// TwinCAT 3 PLC project Tc3UnitTest
// Title: Tc3_UnitTest
// Company: Lorenz Software
// ProjectVersion: 1.0.0.0
// ProgramVersion: 3.1.4026.27
// libraries:
//   Tc2_Standard, * (Beckhoff Automation GmbH)
//   Tc2_System, * (Beckhoff Automation GmbH)
//   Tc2_Utilities, * (Beckhoff Automation GmbH)
// project tree:
//   Framework/Assertions/DataTypes/ AssertionLRealRepresentation.TcDUT, AssertionRealRepresentation.TcDUT
//   Framework/Assertions/GlobalVariables/ Param_Assertions.TcGVL
//   Framework/Assertions/Interfaces/ I_Assertion.TcIO
//   Framework/Assertions/POU/Arrays/Bool/ AssertArrayAllEqual_Bool.TcPOU, AssertArrayContainsArray_Bool.TcPOU, AssertArrayContainsValue_Bool.TcPOU, AssertArrayNoValueChange_Bool.TcPOU, AssertEqualArray_Bool.TcPOU
//   Framework/Assertions/POU/Arrays/Byte/ AssertArrayAllEqual_Byte.TcPOU, AssertArrayContainsArray_Byte.TcPOU, AssertArrayContainsString_Byte.TcPOU, AssertArrayContainsValue_Byte.TcPOU, AssertArrayEndsWithArray_Byte.TcPOU, AssertArrayEndsWithString_Byte.TcPOU, AssertArrayEqualString_Byte.TcPOU, AssertArrayNoValueChange_Byte.TcPOU, AssertArrayStartsWithArray_Byte.TcPOU, AssertArrayStartsWithString_Byte.TcPOU, AssertEqualArray_Byte.TcPOU
//   Framework/Assertions/POU/Arrays/Byte/LengthUntilToken/ AssertLengthUntilArrayEqual_Byte.TcPOU (not stored), AssertLengthUntilArrayGreaterEqual_Byte.TcPOU (not stored), AssertLengthUntilArrayGreaterThan_Byte.TcPOU (not stored), AssertLengthUntilArrayLessEqual_Byte.TcPOU (not stored), AssertLengthUntilArrayLessThan_Byte.TcPOU (not stored), AssertLengthUntilArrayNotEqual_Byte.TcPOU (not stored), AssertLengthUntilValueEqual_Byte.TcPOU (not stored), AssertLengthUntilValueGreaterEqual_Byte.TcPOU (not stored), AssertLengthUntilValueGreaterThan_Byte.TcPOU (not stored), AssertLengthUntilValueLessEqual_Byte.TcPOU (not stored), AssertLengthUntilValueLessThan_Byte.TcPOU (not stored), AssertLengthUntilValueNotEqual_Byte.TcPOU (not stored)
//   Framework/Assertions/POU/Arrays/Byte/TokenCount/ AssertArrayTokenCntEqual_Byte.TcPOU (not stored), AssertArrayTokenCntGreaterEqual_Byte.TcPOU (not stored), AssertArrayTokenCntGreaterThan_Byte.TcPOU (not stored), AssertArrayTokenCntInRange_Byte.TcPOU (not stored), AssertArrayTokenCntLessEqual_Byte.TcPOU (not stored), AssertArrayTokenCntLessThan_Byte.TcPOU (not stored), AssertArrayTokenCntNotEqual_Byte.TcPOU (not stored), AssertArrayTokenCntNotInRange_Byte.TcPOU (not stored), AssertNoArrayToken_Byte.TcPOU (not stored), AssertNoValueToken_Byte.TcPOU (not stored), AssertValueTokenCntEqual_Byte.TcPOU (not stored), AssertValueTokenCntGreaterEqual_Byte.TcPOU (not stored), AssertValueTokenCntGreaterThan_Byte.TcPOU (not stored), AssertValueTokenCntInRange_Byte.TcPOU (not stored), AssertValueTokenCntLessEqual_Byte.TcPOU (not stored), AssertValueTokenCntLessThan_Byte.TcPOU (not stored), AssertValueTokenCntNotEqual_Byte.TcPOU (not stored), AssertValueTokenCntNotInRange_Byte.TcPOU (not stored)
//   Framework/Assertions/POU/Arrays/Char/ AssertArrayAllEqual_Char.TcPOU, AssertArrayContainsArray_Char.TcPOU, AssertArrayContainsString_Char.TcPOU, AssertArrayContainsValue_Char.TcPOU, AssertArrayEndsWithString_Char.TcPOU, AssertArrayEqualString_Char.TcPOU, AssertArrayNoValueChange_Char.TcPOU, AssertArrayStartsWithString_Char.TcPOU, AssertEqualArray_Char.TcPOU
//   Framework/Assertions/POU/Arrays/DInt/ AssertArrayAllEqual_DInt.TcPOU, AssertArrayContainsArray_DInt.TcPOU, AssertArrayContainsValue_DInt.TcPOU, AssertArrayNoValueChange_DInt.TcPOU, AssertEqualArray_DInt.TcPOU
//   Framework/Assertions/POU/Arrays/DWord/ AssertArrayAllEqual_DWord.TcPOU, AssertArrayContainsArray_DWord.TcPOU, AssertArrayContainsValue_DWord.TcPOU, AssertArrayNoValueChange_DWord.TcPOU, AssertEqualArray_DWord.TcPOU
//   Framework/Assertions/POU/Arrays/Int/ AssertArrayAllEqual_Int.TcPOU, AssertArrayContainsArray_Int.TcPOU, AssertArrayContainsValue_Int.TcPOU, AssertArrayNoValueChange_Int.TcPOU, AssertEqualArray_Int.TcPOU
//   Framework/Assertions/POU/Arrays/LInt/ AssertArrayAllEqual_LInt.TcPOU, AssertArrayContainsArray_LInt.TcPOU, AssertArrayContainsValue_LInt.TcPOU, AssertArrayNoValueChange_LInt.TcPOU, AssertEqualArray_LInt.TcPOU
//   Framework/Assertions/POU/Arrays/LReal/ AssertArrayAllElementsFinite_LReal.TcPOU, AssertArrayAllEqual_LReal.TcPOU, AssertArrayContainsArray_LReal.TcPOU, AssertArrayContainsInfinity_LReal.TcPOU, AssertArrayContainsNaN_LReal.TcPOU, AssertArrayContainsNonFinite_LReal.TcPOU, AssertArrayContainsValue_LReal.TcPOU, AssertArrayHasNoInfinity_LReal.TcPOU, AssertArrayHasNoNaN_LReal.TcPOU, AssertArrayNoValueChange_LReal.TcPOU, AssertEqualArray_LReal.TcPOU
//   Framework/Assertions/POU/Arrays/LWord/ AssertArrayAllEqual_LWord.TcPOU, AssertArrayContainsArray_LWord.TcPOU, AssertArrayContainsValue_LWord.TcPOU, AssertArrayNoValueChange_LWord.TcPOU, AssertEqualArray_LWord.TcPOU
//   Framework/Assertions/POU/Arrays/Real/ AssertArrayAllElementsFinite_Real.TcPOU, AssertArrayAllEqual_Real.TcPOU, AssertArrayContainsArray_Real.TcPOU, AssertArrayContainsInfinity_Real.TcPOU, AssertArrayContainsNaN_Real.TcPOU, AssertArrayContainsNonFinite_Real.TcPOU, AssertArrayContainsValue_Real.TcPOU, AssertArrayHasNoInfinity_Real.TcPOU, AssertArrayHasNoNaN_Real.TcPOU, AssertArrayNoValueChange_Real.TcPOU, AssertEqualArray_Real.TcPOU
//   Framework/Assertions/POU/Arrays/SInt/ AssertArrayAllEqual_SInt.TcPOU, AssertArrayContainsArray_SInt.TcPOU, AssertArrayContainsValue_SInt.TcPOU, AssertArrayNoValueChange_SInt.TcPOU, AssertEqualArray_SInt.TcPOU
//   Framework/Assertions/POU/Arrays/UDInt/ AssertArrayAllEqual_UDInt.TcPOU, AssertArrayContainsArray_UDInt.TcPOU, AssertArrayContainsValue_UDInt.TcPOU, AssertArrayNoValueChange_UDInt.TcPOU, AssertEqualArray_UDInt.TcPOU
//   Framework/Assertions/POU/Arrays/UInt/ AssertArrayAllEqual_UInt.TcPOU, AssertArrayContainsArray_UInt.TcPOU, AssertArrayContainsValue_UInt.TcPOU, AssertArrayNoValueChange_UInt.TcPOU, AssertEqualArray_UInt.TcPOU
//   Framework/Assertions/POU/Arrays/ULInt/ AssertArrayAllEqual_ULInt.TcPOU, AssertArrayContainsArray_ULInt.TcPOU, AssertArrayContainsValue_ULInt.TcPOU, AssertArrayNoValueChange_ULInt.TcPOU, AssertEqualArray_ULInt.TcPOU
//   Framework/Assertions/POU/Arrays/USInt/ AssertArrayAllEqual_USInt.TcPOU, AssertArrayContainsArray_USInt.TcPOU, AssertArrayContainsValue_USInt.TcPOU, AssertArrayNoValueChange_USInt.TcPOU, AssertEqualArray_USInt.TcPOU
//   Framework/Assertions/POU/Arrays/WChar/ AssertArrayAllEqual_WChar.TcPOU, AssertArrayContainsArray_WChar.TcPOU, AssertArrayContainsValue_WChar.TcPOU, AssertArrayContainsWString_WChar.TcPOU, AssertArrayEndsWithWString_WChar.TcPOU, AssertArrayEqualWString_WChar.TcPOU, AssertArrayNoValueChange_WChar.TcPOU, AssertArrayStartsWithWString_WChar.TcPOU, AssertEqualArray_WChar.TcPOU
//   Framework/Assertions/POU/Arrays/Word/ AssertArrayAllEqual_Word.TcPOU, AssertArrayContainsArray_Word.TcPOU, AssertArrayContainsValue_Word.TcPOU, AssertArrayContainsWString_Word.TcPOU, AssertArrayEndsWithArray_Word.TcPOU, AssertArrayEndsWithWString_Word.TcPOU, AssertArrayEqualWString_Word.TcPOU, AssertArrayNoValueChange_Word.TcPOU, AssertArrayStartsWithArray_Word.TcPOU, AssertArrayStartsWithWString_Word.TcPOU, AssertEqualArray_Word.TcPOU
//   Framework/Assertions/POU/Arrays/Word/LengthUntilToken/ AssertLengthUntilArrayEqual_Word.TcPOU (not stored), AssertLengthUntilArrayGreaterEqual_Word.TcPOU (not stored), AssertLengthUntilArrayGreaterThan_Word.TcPOU (not stored), AssertLengthUntilArrayLessEqual_Word.TcPOU (not stored), AssertLengthUntilArrayLessThan_Word.TcPOU (not stored), AssertLengthUntilArrayNotEqual_Word.TcPOU (not stored), AssertLengthUntilValueEqual_Word.TcPOU (not stored), AssertLengthUntilValueGreaterEqual_Word.TcPOU (not stored), AssertLengthUntilValueGreaterThan_Word.TcPOU (not stored), AssertLengthUntilValueLessEqual_Word.TcPOU (not stored), AssertLengthUntilValueLessThan_Word.TcPOU (not stored), AssertLengthUntilValueNotEqual_Word.TcPOU (not stored)
//   Framework/Assertions/POU/Arrays/Word/TokenCount/ AssertArrayTokenCntEqual_Word.TcPOU (not stored), AssertArrayTokenCntGreaterEqual_Word.TcPOU (not stored), AssertArrayTokenCntGreaterThan_Word.TcPOU (not stored), AssertArrayTokenCntInRange_Word.TcPOU (not stored), AssertArrayTokenCntLessEqual_Word.TcPOU (not stored), AssertArrayTokenCntLessThan_Word.TcPOU (not stored), AssertArrayTokenCntNotEqual_Word.TcPOU (not stored), AssertArrayTokenCntNotInRange_Word.TcPOU (not stored), AssertNoArrayToken_Word.TcPOU (not stored), AssertNoValueToken_Word.TcPOU (not stored), AssertValueTokenCntEqual_Word.TcPOU (not stored), AssertValueTokenCntGreaterEqual_Word.TcPOU (not stored), AssertValueTokenCntGreaterThan_Word.TcPOU (not stored), AssertValueTokenCntInRange_Word.TcPOU (not stored), AssertValueTokenCntLessEqual_Word.TcPOU (not stored), AssertValueTokenCntLessThan_Word.TcPOU (not stored), AssertValueTokenCntNotEqual_Word.TcPOU (not stored), AssertValueTokenCntNotInRange_Word.TcPOU (not stored)
//   Framework/Assertions/POU/ AssertionBase.TcPOU, AssertionWithEvaluationBase.TcPOU, AssertionEdgeCountBase.TcPOU
//   Framework/Assertions/POU/BasicTypes/Bool/ AssertEqual_Bool.TcPOU, AssertFalse.TcPOU, AssertNotEqual_Bool.TcPOU, AssertNoValueChange_Bool.TcPOU, AssertTrue.TcPOU
//   Framework/Assertions/POU/BasicTypes/Bool/FallingEdge/ AssertFallingEdgeCntEqual.TcPOU (not stored), AssertFallingEdgeCntGreaterEqual.TcPOU (not stored), AssertFallingEdgeCntGreaterThan.TcPOU (not stored), AssertFallingEdgeCntInRange.TcPOU (not stored), AssertFallingEdgeCntLessEqual.TcPOU (not stored), AssertFallingEdgeCntLessThan.TcPOU (not stored), AssertFallingEdgeCntNotEqual.TcPOU (not stored), AssertFallingEdgeCntNotInRange.TcPOU (not stored), AssertNoFallingEdge.TcPOU (not stored)
//   Framework/Assertions/POU/BasicTypes/Bool/RisingEdge/ AssertNoRisingEdge.TcPOU (not stored), AssertRisingEdgeCntEqual.TcPOU (not stored), AssertRisingEdgeCntGreaterEqual.TcPOU (not stored), AssertRisingEdgeCntGreaterThan.TcPOU (not stored), AssertRisingEdgeCntInRange.TcPOU (not stored), AssertRisingEdgeCntLessEqual.TcPOU (not stored), AssertRisingEdgeCntLessThan.TcPOU (not stored), AssertRisingEdgeCntNotEqual.TcPOU (not stored), AssertRisingEdgeCntNotInRange.TcPOU (not stored)
//   Framework/Assertions/POU/BasicTypes/Byte/ AssertContainsBit_Byte.TcPOU, AssertContainsFalse_Byte.TcPOU, AssertContainsTrue_Byte.TcPOU, AssertEqualBit_Byte.TcPOU, AssertEqualMask_Byte.TcPOU, AssertEqual_Byte.TcPOU, AssertFalseBit_Byte.TcPOU, AssertFalseMask_Byte.TcPOU, AssertNotEqualBit_Byte.TcPOU, AssertNotEqualMask_Byte.TcPOU, AssertNotEqual_Byte.TcPOU, AssertNoValueChange_Byte.TcPOU, AssertSequence_Byte.TcPOU, AssertTrueBit_Byte.TcPOU, AssertTrueMask_Byte.TcPOU
//   Framework/Assertions/POU/BasicTypes/Char/ AssertEqual_Char.TcPOU, AssertNotEqual_Char.TcPOU, AssertNoValueChange_Char.TcPOU
//   Framework/Assertions/POU/BasicTypes/Date/ AssertEarlierThan_Date.TcPOU, AssertEqual_Date.TcPOU, AssertInTimespan_Date.TcPOU, AssertLaterThan_Date.TcPOU, AssertNotEqual_Date.TcPOU, AssertNotInTimespan_Date.TcPOU, AssertNoValueChange_Date.TcPOU
//   Framework/Assertions/POU/BasicTypes/DInt/ AssertEqual_DInt.TcPOU, AssertGreaterEqual_DInt.TcPOU, AssertGreaterThan_DInt.TcPOU, AssertInRange_DInt.TcPOU, AssertLessEqual_DInt.TcPOU, AssertLessThan_DInt.TcPOU, AssertNotEqual_DInt.TcPOU, AssertNotInRange_DInt.TcPOU, AssertNoValueChange_DInt.TcPOU, AssertSequence_DInt.TcPOU
//   Framework/Assertions/POU/BasicTypes/DT/ AssertEarlierThan_DT.TcPOU, AssertEqual_DT.TcPOU, AssertInTimespan_DT.TcPOU, AssertLaterThan_DT.TcPOU, AssertNotEqual_DT.TcPOU, AssertNotInTimespan_DT.TcPOU, AssertNoValueChange_DT.TcPOU
//   Framework/Assertions/POU/BasicTypes/DWord/ AssertContainsBit_DWord.TcPOU, AssertContainsFalse_DWord.TcPOU, AssertContainsTrue_DWord.TcPOU, AssertEqualBit_DWord.TcPOU, AssertEqualMask_DWord.TcPOU, AssertEqual_DWord.TcPOU, AssertFalseBit_DWord.TcPOU, AssertFalseMask_DWord.TcPOU, AssertNotEqualBit_DWord.TcPOU, AssertNotEqualMask_DWord.TcPOU, AssertNotEqual_DWord.TcPOU, AssertNoValueChange_DWord.TcPOU, AssertSequence_DWord.TcPOU, AssertTrueBit_DWord.TcPOU, AssertTrueMask_DWord.TcPOU
//   Framework/Assertions/POU/BasicTypes/Int/ AssertEqual_Int.TcPOU, AssertGreaterEqual_Int.TcPOU, AssertGreaterThan_Int.TcPOU, AssertInRange_Int.TcPOU, AssertLessEqual_Int.TcPOU, AssertLessThan_Int.TcPOU, AssertNotEqual_Int.TcPOU, AssertNotInRange_Int.TcPOU, AssertNoValueChange_Int.TcPOU, AssertSequence_Int.TcPOU
//   Framework/Assertions/POU/BasicTypes/LDT/ AssertEarlierThan_LDT.TcPOU, AssertEqual_LDT.TcPOU, AssertInTimespan_LDT.TcPOU, AssertLaterThan_LDT.TcPOU, AssertNotEqual_LDT.TcPOU, AssertNotInTimespan_LDT.TcPOU, AssertNoValueChange_LDT.TcPOU
//   Framework/Assertions/POU/BasicTypes/LInt/ AssertEqual_LInt.TcPOU, AssertGreaterEqual_LInt.TcPOU, AssertGreaterThan_LInt.TcPOU, AssertInRange_LInt.TcPOU, AssertLessEqual_LInt.TcPOU, AssertLessThan_LInt.TcPOU, AssertNotEqual_LInt.TcPOU, AssertNotInRange_LInt.TcPOU, AssertNoValueChange_LInt.TcPOU, AssertSequence_LInt.TcPOU
//   Framework/Assertions/POU/BasicTypes/LReal/ AssertEqualTolerance_LReal.TcPOU, AssertEqual_LReal.TcPOU, AssertGreaterEqual_LReal.TcPOU, AssertGreaterThan_LReal.TcPOU, AssertInRange_LReal.TcPOU, AssertIsFinite_LReal.TcPOU, AssertIsInfinite_LReal.TcPOU, AssertIsNaN_LReal.TcPOU, AssertLessEqual_LReal.TcPOU, AssertLessThan_LReal.TcPOU, AssertNotEqualTolerance_LReal.TcPOU, AssertNotEqual_LReal.TcPOU, AssertNotInRange_LReal.TcPOU, AssertNoValueChange_LReal.TcPOU
//   Framework/Assertions/POU/BasicTypes/LTime/ AssertEarlierThan_LTime.TcPOU, AssertEqual_LTime.TcPOU, AssertInTimespan_LTime.TcPOU, AssertLaterThan_LTime.TcPOU, AssertNotEqual_LTime.TcPOU, AssertNotInTimespan_LTime.TcPOU, AssertNoValueChange_LTime.TcPOU
//   Framework/Assertions/POU/BasicTypes/LTOD/ AssertEarlierThan_LTOD.TcPOU, AssertEqual_LTOD.TcPOU, AssertInTimespan_LTOD.TcPOU, AssertLaterThan_LTOD.TcPOU, AssertNotEqual_LTOD.TcPOU, AssertNotInTimespan_LTOD.TcPOU, AssertNoValueChange_LTOD.TcPOU
//   Framework/Assertions/POU/BasicTypes/LWord/ AssertContainsBit_LWord.TcPOU, AssertContainsFalse_LWord.TcPOU, AssertContainsTrue_LWord.TcPOU, AssertEqualBit_LWord.TcPOU, AssertEqualMask_LWord.TcPOU, AssertEqual_LWord.TcPOU, AssertFalseBit_LWord.TcPOU, AssertFalseMask_LWord.TcPOU, AssertNotEqualBit_LWord.TcPOU, AssertNotEqualMask_LWord.TcPOU, AssertNotEqual_LWord.TcPOU, AssertNoValueChange_LWord.TcPOU, AssertSequence_LWord.TcPOU (not stored), AssertTrueBit_LWord.TcPOU (not stored), AssertTrueMask_LWord.TcPOU (not stored)
//   Framework/Assertions/POU/BasicTypes/Real/ AssertEqualTolerance_Real.TcPOU (not stored), AssertEqual_Real.TcPOU (not stored), AssertGreaterEqual_Real.TcPOU (not stored), AssertGreaterThan_Real.TcPOU (not stored), AssertInRange_Real.TcPOU (not stored), AssertIsFinite_Real.TcPOU (not stored), AssertIsInfinite_Real.TcPOU (not stored), AssertIsNaN_Real.TcPOU (not stored), AssertLessEqual_Real.TcPOU (not stored), AssertLessThan_Real.TcPOU (not stored), AssertNotEqualTolerance_Real.TcPOU (not stored), AssertNotEqual_Real.TcPOU (not stored), AssertNotInRange_Real.TcPOU (not stored), AssertNoValueChange_Real.TcPOU (not stored)
//   Framework/Assertions/POU/BasicTypes/SInt/ AssertEqual_SInt.TcPOU (not stored), AssertGreaterEqual_SInt.TcPOU (not stored), AssertGreaterThan_SInt.TcPOU (not stored), AssertInRange_SInt.TcPOU (not stored), AssertLessEqual_SInt.TcPOU (not stored), AssertLessThan_SInt.TcPOU (not stored), AssertNotEqual_SInt.TcPOU (not stored), AssertNotInRange_SInt.TcPOU (not stored), AssertNoValueChange_SInt.TcPOU (not stored), AssertSequence_SInt.TcPOU (not stored)
//   Framework/Assertions/POU/BasicTypes/String/ AssertContains_String.TcPOU (not stored), AssertEndsWith_String.TcPOU (not stored), AssertEqual_String.TcPOU (not stored), AssertNotEqual_String.TcPOU (not stored), AssertNoValueChange_String.TcPOU (not stored), AssertStartsWith_String.TcPOU (not stored)
//   Framework/Assertions/POU/BasicTypes/Time/ AssertEarlierThan_Time.TcPOU (not stored), AssertEqual_Time.TcPOU (not stored), AssertInTimespan_Time.TcPOU (not stored), AssertLaterThan_Time.TcPOU (not stored), AssertNotEqual_Time.TcPOU (not stored), AssertNotInTimespan_Time.TcPOU (not stored), AssertNoValueChange_Time.TcPOU (not stored)
//   Framework/Assertions/POU/BasicTypes/TOD/ AssertEarlierThan_TOD.TcPOU (not stored), AssertEqual_TOD.TcPOU (not stored), AssertInTimespan_TOD.TcPOU (not stored), AssertLaterThan_TOD.TcPOU (not stored), AssertNotEqual_TOD.TcPOU (not stored), AssertNotInTimespan_TOD.TcPOU (not stored), AssertNoValueChange_TOD.TcPOU (not stored)
//   Framework/Assertions/POU/BasicTypes/UDInt/ AssertEqual_UDInt.TcPOU (not stored), AssertGreaterEqual_UDInt.TcPOU (not stored), AssertGreaterThan_UDInt.TcPOU (not stored), AssertInRange_UDInt.TcPOU (not stored), AssertLessEqual_UDInt.TcPOU (not stored), AssertLessThan_UDInt.TcPOU (not stored), AssertNotEqual_UDInt.TcPOU (not stored), AssertNotInRange_UDInt.TcPOU (not stored), AssertNoValueChange_UDInt.TcPOU (not stored), AssertSequence_UDInt.TcPOU (not stored)
//   Framework/Assertions/POU/BasicTypes/UInt/ AssertEqual_UInt.TcPOU (not stored), AssertGreaterEqual_UInt.TcPOU (not stored), AssertGreaterThan_UInt.TcPOU (not stored), AssertInRange_UInt.TcPOU (not stored), AssertLessEqual_UInt.TcPOU (not stored), AssertLessThan_UInt.TcPOU (not stored), AssertNotEqual_UInt.TcPOU (not stored), AssertNotInRange_UInt.TcPOU (not stored), AssertNoValueChange_UInt.TcPOU (not stored), AssertSequence_UInt.TcPOU (not stored)
//   Framework/Assertions/POU/BasicTypes/ULInt/ AssertEqual_ULInt.TcPOU (not stored), AssertGreaterEqual_ULInt.TcPOU (not stored), AssertGreaterThan_ULInt.TcPOU (not stored), AssertInRange_ULInt.TcPOU (not stored), AssertLessEqual_ULInt.TcPOU (not stored), AssertLessThan_ULInt.TcPOU (not stored), AssertNotEqual_ULInt.TcPOU (not stored), AssertNotInRange_ULInt.TcPOU (not stored), AssertNoValueChange_ULInt.TcPOU (not stored), AssertSequence_ULInt.TcPOU (not stored)
//   Framework/Assertions/POU/BasicTypes/USInt/ AssertEqual_USInt.TcPOU (not stored), AssertGreaterEqual_USInt.TcPOU (not stored), AssertGreaterThan_USInt.TcPOU (not stored), AssertInRange_USInt.TcPOU (not stored), AssertLessEqual_USInt.TcPOU (not stored), AssertLessThan_USInt.TcPOU (not stored), AssertNotEqual_USInt.TcPOU (not stored), AssertNotInRange_USInt.TcPOU (not stored), AssertNoValueChange_USInt.TcPOU (not stored), AssertSequence_USInt.TcPOU (not stored)
//   Framework/Assertions/POU/BasicTypes/WChar/ AssertEqual_WChar.TcPOU (not stored), AssertNotEqual_WChar.TcPOU (not stored), AssertNoValueChange_WChar.TcPOU (not stored)
//   Framework/Assertions/POU/BasicTypes/Word/ AssertContainsBit_Word.TcPOU (not stored), AssertContainsFalse_Word.TcPOU (not stored), AssertContainsTrue_Word.TcPOU (not stored), AssertEqualBit_Word.TcPOU (not stored), AssertEqualMask_Word.TcPOU (not stored), AssertEqual_Word.TcPOU (not stored), AssertFalseBit_Word.TcPOU (not stored), AssertFalseMask_Word.TcPOU (not stored), AssertNotEqualBit_Word.TcPOU (not stored), AssertNotEqualMask_Word.TcPOU (not stored), AssertNotEqual_Word.TcPOU (not stored), AssertNoValueChange_Word.TcPOU (not stored), AssertSequence_Word.TcPOU (not stored), AssertTrueBit_Word.TcPOU (not stored), AssertTrueMask_Word.TcPOU (not stored)
//   Framework/Assertions/POU/BasicTypes/WString/ AssertContains_WString.TcPOU (not stored), AssertEndsWith_WString.TcPOU (not stored), AssertEqual_WString.TcPOU (not stored), AssertNotEqual_WString.TcPOU (not stored), AssertNoValueChange_WString.TcPOU (not stored), AssertStartsWith_WString.TcPOU (not stored)
//   Framework/Assertions/POU/Utilities/ CountArrayTokens_Byte.TcPOU, CountArrayTokens_Word.TcPOU, CountValueTokens_Byte.TcPOU, CountValueTokens_Word.TcPOU, CreateAssertionTextValue_BinaryFloat.TcPOU, CreateAssertionTextValue_ByteArray.TcPOU, CreateAssertionTextValue_Char.TcPOU, CreateAssertionTextValue_Hex.TcPOU, CreateAssertionTextValue_LReal.TcPOU, CreateAssertionTextValue_Real.TcPOU, CreateAssertionTextValue_String.TcPOU, CreateAssertionTextValue_WChar.TcPOU, CreateAssertionTextValue_WordArray.TcPOU, CreateAssertionTextValue_WString.TcPOU, DateToDayNumber.TcPOU, FindArrayToken_Byte.TcPOU, FindArrayToken_Word.TcPOU, FindValueToken_Byte.TcPOU, FindValueToken_Word.TcPOU, IsAssertionStringLengthValid.TcPOU, IsAssertionWStringLengthValid.TcPOU, IsTimeOfDayValid_LTOD.TcPOU, IsTimeOfDayValid_TOD.TcPOU, IsWithinTolerance_LReal.TcPOU, IsWithinTolerance_Real.TcPOU, TextContains_String.TcPOU, TextContains_WString.TcPOU, TextEndsWith_String.TcPOU, TextStartsWith_String.TcPOU, TextEndsWith_WString.TcPOU, TextStartsWith_WString.TcPOU
//   Framework/Common/DataTypes/ E_ExecutionStatus.TcDUT, E_OrchestrationMode.TcDUT, E_OrchestratorTask.TcDUT, E_Result.TcDUT, E_State.TcDUT, ST_Command.TcDUT, ST_ContractInfo.TcDUT, ST_ExecutionStatus.TcDUT
//   Framework/Common/Fifo/DataTypes/ E_FifoResult.TcDUT, ST_FifoStatus.TcDUT
//   Framework/Common/Fifo/POU/ Fifo.TcPOU
//   Framework/Common/GlobalVariables/ Global_Version.TcGVL, GVL_Constants.TcGVL, GVL_UnitTest.TcGVL
//   Framework/Common/Interfaces/ I_Orchestratable.TcIO, I_OrchestratableCollection.TcIO, I_Orchestrator.TcIO, I_ResultAggregator.TcIO, I_ResultProvider.TcIO
//   Framework/Common/POU/ Stopwatch.TcPOU, GetFrameworkVersion.TcPOU, IsNameValid.TcPOU, Orchestrator.TcPOU, ResultAggregator.TcPOU
//   Framework/EventBuffer/DataTypes/ E_EventPublishResult.TcDUT, E_EventReservationResult.TcDUT, E_EventSeverity.TcDUT, E_EventType.TcDUT, E_OwnerScope.TcDUT, ST_Event.TcDUT, ST_EventBufferCommand.TcDUT, ST_EventBufferStatus.TcDUT, ST_EventStream.TcDUT
//   Framework/EventBuffer/GlobalVariables/ GVL_EventBuffer.TcGVL, Param_EventBuffer.TcGVL
//   Framework/EventBuffer/Interfaces/ I_EventBuffer.TcIO, I_EventPublisher.TcIO
//   Framework/EventBuffer/POU/AggregationEvents/ CreateRunAggregationEvent.TcPOU, CreateTestCaseAggregationEvent.TcPOU, CreateTestSuiteAggregationEvent.TcPOU
//   Framework/EventBuffer/POU/ EventBuffer.TcPOU, EventBufferDiagConsumer.TcPOU
//   Framework/EventBuffer/POU/FrameworkEvents/ CreateFrameworkEvent.TcPOU, CreateInvalidStateTransitionEvent.TcPOU, CreateResetWarningEvent.TcPOU
//   Framework/EventBuffer/POU/ResultEvents/ CreateAssertionErrorEvent.TcPOU, CreateAssertionFailedEvent.TcPOU, CreateResultEvent.TcPOU
//   Framework/EventBuffer/POU/StateTransitionEvents/ CreateStateTransitionEvent.TcPOU, CreateTestCaseOrchestratorStateTransitionEvent.TcPOU, CreateTestSuiteOrchestratorStateTransitionEvent.TcPOU
//   Framework/EventBuffer/POU/TriggerEvents/ CreateAbortEvent.TcPOU, CreateResetEvent.TcPOU, CreateStartEvent.TcPOU
//   Framework/EventBuffer/POU/Utilities/ SelectResultSeverity.TcPOU
//   Framework/Preparation/DataTypes/ ST_PreparationStatus.TcDUT
//   Framework/Preparation/Interfaces/ I_Preparation.TcIO
//   Framework/Preparation/POU/ PreparationBase.TcPOU, PreparationMock.TcPOU
//   Framework/RunControl/DataTypes/ ST_RunConfig.TcDUT, ST_RunControl.TcDUT, ST_RunControlCommunication.TcDUT, ST_RunControlStatus.TcDUT, ST_TestSuiteCollectionConfig.TcDUT
//   Framework/RunControl/Interfaces/ I_RunControl.TcIO
//   Framework/RunControl/POU/ RunControlBase.TcPOU, RunControlCommandAdapter.TcPOU, RunControlConfigurationBuilder.TcPOU
//   Framework/TestCases/DataTypes/ ST_TestCaseConfig.TcDUT, ST_TestCaseExecutionStatus.TcDUT, ST_TestCaseStatus.TcDUT
//   Framework/TestCases/Interfaces/ I_TestCase.TcIO
//   Framework/TestCases/POU/ TestCaseBase.TcPOU, TestCaseMock.TcPOU
//   Framework/TestSuites/DataTypes/ ST_TestCaseCollectionConfig.TcDUT, ST_TestSuiteConfig.TcDUT, ST_TestSuiteStatus.TcDUT
//   Framework/TestSuites/Interfaces/ I_TestSuite.TcIO
//   Framework/TestSuites/POU/ TestSuiteBase.TcPOU, TestSuiteConfigurationBuilder.TcPOU, TestSuiteMock.TcPOU
//   Runtime/ PlcTask.TcTTO, MAIN.TcPOU
//   SelfTests/Helper/Orchestration/DataTypes/ E_OrchestrationArrayLayout.TcDUT, ST_OrchestrationCalls.TcDUT, ST_OrchestrationCycle.TcDUT, ST_OrchestrationObservation.TcDUT, ST_OrchestrationStep.TcDUT
//   SelfTests/Helper/Orchestration/ OrchestrationChildDouble.TcPOU, OrchestrationCollectionDouble.TcPOU, OrchestratorProbe.TcPOU, OrchestrationTestBase.TcPOU
//   SelfTests/RunControl/ RunControl.TcPOU
//   SelfTests/TestCases/TestSuite_AssertionArrays/ Test_AssertionArrayComparison.TcPOU, Test_AssertionArrayPatternSearch.TcPOU, Test_AssertionArrayTextBridge.TcPOU, Test_AssertionArrayValueSearch.TcPOU, Test_AssertionFloatingPointArray.TcPOU, Test_AssertionMaskedArrayComparison.TcPOU
//   SelfTests/TestCases/TestSuite_AssertionComparisons/ Test_AssertionBitEquality.TcPOU, Test_AssertionBooleanComparisons.TcPOU, Test_AssertionCharacterEquality.TcPOU, Test_AssertionDateNormalization.TcPOU, Test_AssertionDurationComparisons.TcPOU, Test_AssertionLTODDomain.TcPOU, Test_AssertionScalarDiagnostics.TcPOU, Test_AssertionSignedRanges.TcPOU, Test_AssertionSignedRelations.TcPOU, Test_AssertionTODDomain.TcPOU, Test_AssertionUnsignedRanges.TcPOU, Test_AssertionUnsignedRelations.TcPOU
//   SelfTests/TestCases/TestSuite_AssertionFloatingPoint/DataTypes/ FloatingPointBits_LReal.TcDUT, FloatingPointBits_Real.TcDUT
//   SelfTests/TestCases/TestSuite_AssertionFloatingPoint/ Test_AssertionArrayClassification_LReal.TcPOU, Test_AssertionArrayClassification_Real.TcPOU, Test_AssertionClassification_LReal.TcPOU, Test_AssertionClassification_Real.TcPOU, Test_AssertionFiniteBoundaries_LReal.TcPOU, Test_AssertionFiniteBoundaries_Real.TcPOU, Test_AssertionNonFinite_LReal.TcPOU, Test_AssertionNonFinite_Real.TcPOU, Test_AssertionRelations_LReal.TcPOU, Test_AssertionRelations_Real.TcPOU, Test_AssertionTolerance_LReal.TcPOU, Test_AssertionTolerance_Real.TcPOU
//   SelfTests/TestCases/TestSuite_AssertionLifecycle/Helper/ AssertionEvaluationSubject.TcPOU, AssertionLifecycleSubject.TcPOU, AssertionParentIdentity.TcPOU
//   SelfTests/TestCases/TestSuite_AssertionLifecycle/ Test_AssertionActivity.TcPOU, Test_AssertionEscalation.TcPOU, Test_AssertionInitialization.TcPOU, Test_AssertionResetReuse.TcPOU, Test_AssertionUninitialized.TcPOU
//   SelfTests/TestCases/TestSuite_AssertionObservation/ Test_AssertionArraySnapshot.TcPOU, Test_AssertionEdgeCount.TcPOU, Test_AssertionEdgeObservation.TcPOU, Test_AssertionFloatingSnapshot.TcPOU, Test_AssertionScalarObservation.TcPOU, Test_AssertionSequence.TcPOU
//   SelfTests/TestCases/TestSuite_AssertionText/ Test_AssertionArrayTokenCount.TcPOU, Test_AssertionLengthUntil.TcPOU, Test_AssertionTextComparison.TcPOU, Test_AssertionTextDiagnostics.TcPOU, Test_AssertionTextSearch.TcPOU, Test_AssertionValueTokenCount.TcPOU
//   SelfTests/TestCases/TestSuite_AssertionVariants/ Test_AssertionBitSelection.TcPOU, Test_AssertionCountPredicates.TcPOU, Test_AssertionMaskPredicates.TcPOU, Test_AssertionNarrowIntegers.TcPOU, Test_AssertionTemporalVariants.TcPOU
//   SelfTests/TestCases/TestSuite_CommandAdapter/DataTypes/ E_AdapterCommand.TcDUT
//   SelfTests/TestCases/TestSuite_CommandAdapter/Helper/ RunControlRequestRecorder.TcPOU
//   SelfTests/TestCases/TestSuite_CommandAdapter/ Test_CommandAdapterInitialization.TcPOU, Test_CommandIndependence.TcPOU, Test_CommandQualification.TcPOU
//   SelfTests/TestCases/TestSuite_EventBufferReset/Helper/ ActiveResetBufferProbe.TcPOU, BufferCommandProbe.TcPOU, BufferReleaseSuiteDouble.TcPOU, BufferResetRunControlProbe.TcPOU
//   SelfTests/TestCases/TestSuite_EventBufferReset/ Test_BufferResetActiveRun.TcPOU, Test_BufferResetCommands.TcPOU, Test_BufferResetEpochs.TcPOU
//   SelfTests/TestCases/TestSuite_EventDelivery/ Test_EventBufferFull.TcPOU, Test_EventContent.TcPOU, Test_EventDeleteCommandBoundary.TcPOU, Test_EventDeleteLostSequence.TcPOU, Test_EventDeleteWatermarks.TcPOU, Test_EventDeleteWrappedFull.TcPOU, Test_EventRingOrder.TcPOU, Test_EventStorageBinding.TcPOU
//   SelfTests/TestCases/TestSuite_EventReservation/Helper/ ReservationChildProbe.TcPOU, ReservationResetChild.TcPOU, ReservationSuiteProbe.TcPOU
//   SelfTests/TestCases/TestSuite_EventReservation/ Test_ActiveReservationLoss.TcPOU, Test_ExecutionReservationAccounting.TcPOU, Test_HierarchicalReservationRelease.TcPOU, Test_ImpossibleExecutionBudget.TcPOU, Test_ImpossibleResetBudget.TcPOU, Test_LateResetReservationRelease.TcPOU, Test_ReservationAdmission.TcPOU, Test_ResetReservationAccounting.TcPOU
//   SelfTests/TestCases/TestSuite_Orchestrator/ Test_OrchestratorExecutionBudgetError.TcPOU, Test_OrchestratorExecutionCapacityWait.TcPOU, Test_OrchestratorResetCapacityWait.TcPOU, Test_OrchestratorShiftedBounds.TcPOU, Test_OrchestratorNegativeBounds.TcPOU, Test_OrchestratorUnusedCapacity.TcPOU, Test_OrchestratorSingleChild.TcPOU, Test_OrchestratorIdleReadiness.TcPOU, Test_OrchestratorMissingStartReaction.TcPOU, Test_OrchestratorChildError.TcPOU, Test_OrchestratorUnexpectedAbort.TcPOU, Test_OrchestratorAbortInterruption.TcPOU, Test_OrchestratorIdleInterruption.TcPOU, Test_OrchestratorResetInterruption.TcPOU, Test_OrchestratorResetContinuesAfterError.TcPOU, Test_OrchestratorRepeatAfterReset.TcPOU
//   SelfTests/TestCases/TestSuite_ParallelOrchestration/ Test_ParallelAbortMixedProgress.TcPOU, Test_ParallelChildError.TcPOU, Test_ParallelFailedResultContinues.TcPOU, Test_ParallelFirstFittingAdmission.TcPOU, Test_ParallelMissingStartReaction.TcPOU, Test_ParallelReadinessLost.TcPOU, Test_ParallelResetOverlappingExecution.TcPOU, Test_ParallelUnequalDurations.TcPOU
//   SelfTests/TestCases/TestSuite_ParallelSlotsOrchestration/ Test_SlotsAbortAtBoundary.TcPOU, Test_SlotsFinalGroupCompletion.TcPOU, Test_SlotsFirstFittingAdmission.TcPOU, Test_SlotsMissingStartReaction.TcPOU, Test_SlotsNextSlotReadinessLost.TcPOU, Test_SlotsWaitForGroupCompletion.TcPOU
//   SelfTests/TestCases/TestSuite_Preparation/Helper/ PreparationResource.TcPOU, PreparationStatusProbe.TcPOU, Prepare_ValueAtTarget.TcPOU, Prepare_ZeroViaOne.TcPOU
//   SelfTests/TestCases/TestSuite_Preparation/ Test_PreparationCompletionTracksTarget.TcPOU, Test_PreparationDisableAndReenable.TcPOU, Test_PreparationDisabledObservation.TcPOU, Test_PreparationInitialStatus.TcPOU, Test_PreparationMockInputs.TcPOU, Test_PreparationReachesTarget.TcPOU, Test_PreparationResourceError.TcPOU, Test_PreparationStatusProjection.TcPOU
//   SelfTests/TestCases/TestSuite_RunControlConfigurationBuilder/ Test_RunControlBuilderCapacity.TcPOU, Test_RunControlBuilderFinalizeReuse.TcPOU, Test_RunControlBuilderParallel.TcPOU, Test_RunControlBuilderRegistrationErrors.TcPOU, Test_RunControlBuilderSerial.TcPOU, Test_RunControlBuilderSlotInsertion.TcPOU
//   SelfTests/TestCases/TestSuite_RunControlLifecycle/DataTypes/ E_RunControlCompletionScenario.TcDUT, E_RunControlLifecycleScenario.TcDUT
//   SelfTests/TestCases/TestSuite_RunControlLifecycle/Helper/ RunControlIntegrationSubject.TcPOU, RunControlLifecycleProbe.TcPOU, RunControlSuiteDouble.TcPOU
//   SelfTests/TestCases/TestSuite_RunControlLifecycle/ Test_RunControlCompletion.TcPOU, Test_RunControlExceptionalLifecycle.TcPOU, Test_RunControlInitialization.TcPOU, Test_RunControlNormalLifecycle.TcPOU, Test_RunControlRealComposition.TcPOU, Test_RunControlRequests.TcPOU, Test_RunControlTaskMapping.TcPOU
//   SelfTests/TestCases/TestSuite_SerialOrchestration/ Test_SerialFailedResultContinues.TcPOU, Test_SerialImmediateCompletion.TcPOU, Test_SerialNotReadyCandidate.TcPOU, Test_SerialRegistrationOrder.TcPOU, Test_SerialUnequalDurations.TcPOU
//   SelfTests/TestCases/TestSuite_Smoke/ Test_Smoke.TcPOU
//   SelfTests/TestCases/TestSuite_TestCaseLifecycle/Helper/DataTypes/ E_LifecycleHook.TcDUT (not stored), ST_LifecycleHook.TcDUT (not stored), ST_LifecycleStep.TcDUT (not stored)
//   SelfTests/TestCases/TestSuite_TestCaseLifecycle/Helper/ TestCaseInitializationProbe.TcPOU, TestCaseLifecycleProbe.TcPOU, TestCaseLifecycleTestBase.TcPOU
//   SelfTests/TestCases/TestSuite_TestCaseLifecycle/ Test_LifecycleAbort.TcPOU, Test_LifecycleAbortError.TcPOU, Test_LifecycleAbortTimeout.TcPOU, Test_LifecycleAlreadyPrepared.TcPOU, Test_LifecycleExecutionTimeout.TcPOU, Test_LifecycleFailedResult.TcPOU, Test_LifecycleFailedToError.TcPOU, Test_LifecycleInitialization.TcPOU, Test_LifecycleInvalidPreparationTransition.TcPOU, Test_LifecycleInvalidTestAdvance.TcPOU, Test_LifecycleMultipleStates.TcPOU, Test_LifecyclePreparationError.TcPOU, Test_LifecyclePreparationTimeout.TcPOU, Test_LifecycleRepeatAfterAbort.TcPOU, Test_LifecycleRepeatAfterError.TcPOU, Test_LifecycleRepeatAfterFailed.TcPOU, Test_LifecycleRepeatAfterPassed.TcPOU, Test_LifecycleResetDuringExecution.TcPOU, Test_LifecycleResetError.TcPOU, Test_LifecycleResetTimeout.TcPOU, Test_LifecycleSinglePreparation.TcPOU, Test_LifecycleWithoutPreparation.TcPOU
//   SelfTests/TestCases/TestSuite_TestSuiteConfigurationBuilder/ Test_SuiteBuilderCapacity.TcPOU, Test_SuiteBuilderFinalizeReuse.TcPOU, Test_SuiteBuilderParallel.TcPOU, Test_SuiteBuilderRegistrationErrors.TcPOU, Test_SuiteBuilderSerial.TcPOU, Test_SuiteBuilderSlotInsertion.TcPOU
//   SelfTests/TestCases/TestSuite_TestSuiteLifecycle/DataTypes/ E_SuiteLifecycleScenario.TcDUT
//   SelfTests/TestCases/TestSuite_TestSuiteLifecycle/Helper/ SuiteIntegrationChild.TcPOU, SuiteIntegrationSubject.TcPOU, SuiteLifecycleChildDouble.TcPOU, SuiteOrchestratorDouble.TcPOU, TestSuiteLifecycleProbe.TcPOU, TestSuiteMockProbe.TcPOU
//   SelfTests/TestCases/TestSuite_TestSuiteLifecycle/ Test_SuiteExceptionalLifecycle.TcPOU, Test_SuiteFinalization.TcPOU, Test_SuiteInitialization.TcPOU, Test_SuiteMockRepeatedReset.TcPOU, Test_SuiteNormalLifecycle.TcPOU, Test_SuiteReadiness.TcPOU, Test_SuiteRealComposition.TcPOU, Test_SuiteReservationRelease.TcPOU
//   SelfTests/TestSuites/ TestSuite_AssertionArrays.TcPOU, TestSuite_AssertionComparisons.TcPOU, TestSuite_AssertionFloatingPoint.TcPOU, TestSuite_AssertionLifecycle.TcPOU, TestSuite_AssertionObservation.TcPOU, TestSuite_AssertionText.TcPOU, TestSuite_AssertionVariants.TcPOU, TestSuite_CommandAdapter.TcPOU, TestSuite_EventBufferReset.TcPOU, TestSuite_EventDelivery.TcPOU, TestSuite_EventReservation.TcPOU, TestSuite_Orchestrator.TcPOU, TestSuite_ParallelOrchestration.TcPOU, TestSuite_ParallelSlotsOrchestration.TcPOU, TestSuite_Preparation.TcPOU, TestSuite_RunControlConfigurationBuilder.TcPOU, TestSuite_RunControlLifecycle.TcPOU, TestSuite_SerialOrchestration.TcPOU, TestSuite_Smoke.TcPOU, TestSuite_TestCaseLifecycle.TcPOU, TestSuite_TestSuiteConfigurationBuilder.TcPOU, TestSuite_TestSuiteLifecycle.TcPOU
// real-time tasks:
//   TASK PlcTask: cycle T#1ms, priority 20, ADS port 350

CONFIGURATION Tc3UnitTest
    RESOURCE PLC ON TwinCAT3
        TASK PlcTask(INTERVAL := T#1ms, PRIORITY := 20);
        PROGRAM MAIN WITH PlcTask : MAIN;
    END_RESOURCE
END_CONFIGURATION

// ---- Framework/Assertions/DataTypes/AssertionLRealRepresentation.TcDUT
{region 'Documentation'}
(*!
<summary>Internal IEEE binary64 view for diagnostic formatting without floating-point operations.</summary>
*)
{endregion}
TYPE INTERNAL AssertionLRealRepresentation :
UNION
    Value : LREAL; //! Floating-point view of the shared 64-bit storage.
    Bits : LWORD; //! Raw IEEE binary64 bit pattern of the same storage.
END_UNION
END_TYPE

// ---- Framework/Assertions/DataTypes/AssertionRealRepresentation.TcDUT
{region 'Documentation'}
(*!
<summary>Internal IEEE binary32 view for diagnostic formatting without floating-point operations.</summary>
*)
{endregion}
TYPE INTERNAL AssertionRealRepresentation :
UNION
    Value : REAL; //! Floating-point view of the shared 32-bit storage.
    Bits : DWORD; //! Raw IEEE binary32 bit pattern of the same storage.
END_UNION
END_TYPE

// ---- Framework/Common/DataTypes/E_ExecutionStatus.TcDUT
{region 'Documentation'}
(*!
<summary>Coarse execution classification derived from the owner state.</summary>
*)
{endregion}
{attribute 'qualified_only'}
{attribute 'strict'}
TYPE E_ExecutionStatus :
(
    Error := -10, //! Execution cannot continue normally.
    Unknown := 0, //! No classified observation is available.
    Inactive := 1, //! Inactive execution classification retained by the contract.
    NotReady := 9, //! Not ready to begin execution.
    Idle := 10, //! Reset-defined idle execution condition.
    Starting := 20, //! Start processing is in progress.
    Running := 30, //! Execution is active.
    Completing := 40, //! Finalization is in progress.
    Completed := 50, //! Execution has ended; inspect Result for its outcome.
    Aborting := 60, //! Controlled termination is in progress.
    Aborted := 70, //! Legacy value; not used as a stable final status by new owner logic.
    Reset := 80 //! Reset processing is in progress.
) INT := Unknown;
END_TYPE

// ---- Framework/Common/DataTypes/E_OrchestrationMode.TcDUT
{region 'Documentation'}
(*!
<summary>Child scheduling strategy represented by effective execution slots.</summary>
*)
{endregion}
{attribute 'qualified_only'}
{attribute 'strict'}
TYPE E_OrchestrationMode :
(
    Serial := 0, //! Run one child per slot, in registration order.
    Parallel := 1, //! Run all children in one shared slot.
    ParallelSlots := 2 //! Run children in ascending explicit slots; finish one slot before starting the next.
);
END_TYPE

// ---- Framework/Common/DataTypes/E_OrchestratorTask.TcDUT
{region 'Documentation'}
(*!
<summary>Owner-requested orchestration work; independent of the owner lifecycle.</summary>
*)
{endregion}
{attribute 'qualified_only'}
{attribute 'strict'}
TYPE E_OrchestratorTask :
(
    Idle := 0, //! No new child work is dispatched.
    Reset := 1, //! Dispatch capacity-admitted child resets and observe their completion.
    Execution := 2, //! Dispatch capacity-admitted starts by slot and observe completion.
    Abort := 3 //! Request and observe controlled termination of active children.
);
END_TYPE

// ---- Framework/Common/DataTypes/E_Result.TcDUT
{region 'Documentation'}
(*!
<summary>Stable evaluation result; numeric order is not severity order.</summary>
*)
{endregion}
{attribute 'qualified_only'}
{attribute 'strict'}
TYPE E_Result :
(
    Error := -10, //! Execution or evaluation error; highest result severity.
    NotEvaluated := 0, //! No evaluated outcome; neutral result after reset.
    Passed := 10, //! Evaluated checks succeeded.
    // SA0027: Qualified enum member; retained despite the analyzer's name-collision report.
    {attribute 'analysis' := '-27'}
    Failed := 20, //! An evaluated check failed; lower severity than Abort or Error.
    Abort := 30 //! Execution aborted; lower severity than Error, higher than Failed.
) INT := NotEvaluated;
END_TYPE

// ---- Framework/Common/DataTypes/E_State.TcDUT
{region 'Documentation'}
(*!
<summary>Owner lifecycle state. Non-strict for configured Preparation and Test state intervals.</summary>
*)
{endregion}
{attribute 'qualified_only'}
TYPE E_State :
(
    Error := -10, //! Error state value; active errors use controlled error finalization.
    Uninitialized := 0, //! Not yet in a reset-defined executable state.
    Reset := 1, //! Reset work in progress.
    Idle := 10, //! Reset-defined base state; readiness is reported separately.
    Starting := 11, //! Start accepted; execution setup in progress.
    Preparing := 20, //! First configured Preparation state; subsequent values precede Running.
    Running := 50, //! First configured Test state, or active Suite/Run execution.
    Completing := 80, //! Finalization phase before stable completion.
    Completed := 89, //! Stable terminal state; result determines the outcome.
    Aborting := 90, //! Controlled termination requested by Abort.
    AbortingFromError := 91, //! Controlled termination caused by an execution error.
    Aborted := 99 //! Legacy aborted state; new owners finalize in Completed.
) INT := Uninitialized;
END_TYPE

// ---- Framework/Common/DataTypes/ST_Command.TcDUT
{region 'Documentation'}
(*!
<summary>Lifecycle request flags; external qualification and clearing belong to the command adapter.</summary>
*)
{endregion}
TYPE ST_Command :
STRUCT
    {attribute 'OPC.UA.DA.Access' := '3'}
    Start : BOOL := FALSE; //! External one-shot Start request, qualified and cleared by the command adapter.
    {attribute 'OPC.UA.DA.Access' := '3'}
    Abort : BOOL := FALSE; //! External one-shot Abort request for active execution, qualified and cleared by the command adapter.
    {attribute 'OPC.UA.DA.Access' := '3'}
    Reset : BOOL := FALSE; //! External one-shot lifecycle Reset request, qualified and cleared by the command adapter.
END_STRUCT
END_TYPE

// ---- Framework/Common/DataTypes/ST_ContractInfo.TcDUT
{region 'Documentation'}
(*!
<summary>Compatibility and effective library-version metadata.</summary>
*)
{endregion}
TYPE ST_ContractInfo :
STRUCT
    {attribute 'OPC.UA.DA.Access' := '1'}
    ContractVersion : STRING(GVL_Constants.VersionLength) := ''; //! Version of this communication contract, formatted as Major.Minor.Build.
    {attribute 'OPC.UA.DA.Access' := '1'}
    FrameworkVersion : STRING(GVL_Constants.VersionLength) := ''; //! Effective library version as Major.Minor.Build; TwinCAT revision is omitted.
END_STRUCT
END_TYPE

// ---- Framework/Common/DataTypes/ST_ExecutionStatus.TcDUT
{region 'Documentation'}
(*!
<summary>Owner execution and result snapshot.</summary>
*)
{endregion}
TYPE ST_ExecutionStatus :
STRUCT
    {attribute 'OPC.UA.DA.Access' := '1'}
    State : E_State := E_State.Uninitialized; //! Owner's detailed lifecycle state, including configured Test Case phases.
    {attribute 'OPC.UA.DA.Access' := '1'}
    ExecutionStatus : E_ExecutionStatus := E_ExecutionStatus.Unknown; //! Coarse execution classification derived from State.
    {attribute 'OPC.UA.DA.Access' := '1'}
    Result : E_Result := E_Result.NotEvaluated; //! Current held evaluation result; numeric order is not severity order.
    {attribute 'OPC.UA.DA.Access' := '1'}
    Uninitialized : BOOL := FALSE; //! Owner has not reached a reset-defined executable base state.
    {attribute 'OPC.UA.DA.Access' := '1'}
    ConfigError : BOOL := FALSE; //! Owner setup is invalid or has not yet been validated.
    {attribute 'OPC.UA.DA.Access' := '1'}
    Ready : BOOL := FALSE; //! Owner is initialized, Idle and ready to accept Start.
    {attribute 'OPC.UA.DA.Access' := '1'}
    Running : BOOL := FALSE; //! Owner is in its active execution phase.
    {attribute 'OPC.UA.DA.Access' := '1'}
    Completed : BOOL := FALSE; //! Owner has reached its terminal Completed state; does not imply Passed.
    {attribute 'OPC.UA.DA.Access' := '1'}
    Aborted : BOOL := FALSE; //! Owner completed with Abort result.
    {attribute 'OPC.UA.DA.Access' := '1'}
    // SA0033: Contract status field retained even when not consumed by this application.
    {attribute 'analysis' := '-33'}
    Inactive : BOOL := FALSE; //! Contract-reserved inactive indication; retained for compatible consumers.
    {attribute 'OPC.UA.DA.Access' := '1'}
    Error : BOOL := FALSE; //! Owner reports an error, including Result = Error.
END_STRUCT
END_TYPE

// ---- Framework/Common/Fifo/DataTypes/E_FifoResult.TcDUT
{region 'Documentation'}
(*!
<summary>Internal FIFO operation results; positive transfer slots are returned separately from these zero or negative outcomes.</summary>
*)
{endregion}
{attribute 'qualified_only'}
TYPE INTERNAL E_FifoResult :
(
    NoTransfer := 0, //! No event transferred, for example an empty read or full insertion.
    ConfigError := -1, //! Storage configuration or retained binding is invalid.
    IndexError := -2, //! Stored ring indices are invalid.
    DataError := -3, //! Data access would violate the storage requirements.
    ReleaseCountError := -4 //! Requested release count exceeds the queued event count.
) INT;
END_TYPE

// ---- Framework/Common/Fifo/DataTypes/ST_FifoStatus.TcDUT
{region 'Documentation'}
(*!
<summary>FIFO binding, logical ring indices and derived occupancy snapshot; payload storage remains caller-owned.</summary>
*)
{endregion}
TYPE ST_FifoStatus :
STRUCT
    {attribute 'OPC.UA.DA.Access' := '1'}
    IndexIn : UINT; //! One-based next write position; equal to IndexOut when the ring is empty.
    {attribute 'OPC.UA.DA.Access' := '1'}
    IndexOut : UINT; //! One-based oldest occupied position; read from here before acknowledging events.
    {attribute 'OPC.UA.DA.Access' := '1'}
    ConfigError : BOOL; //! Storage is uninitialized or its binding/configuration is invalid.
    {attribute 'OPC.UA.DA.Access' := '1'}
    IndexError : BOOL; //! At least one stored ring index is outside the configured range.
    {attribute 'OPC.UA.DA.Access' := '1'}
    BufferAlmostFull : BOOL; //! Exactly one usable event slot remains free.
    {attribute 'OPC.UA.DA.Access' := '1'}
    BufferFull : BOOL; //! No usable event slot remains; the physical ring always retains one unused position.
    {attribute 'OPC.UA.DA.Access' := '1'}
    BufferEmpty : BOOL; //! No event is currently queued.
    {attribute 'OPC.UA.DA.Access' := '1'}
    ElementCount : UINT; //! Number of queued events, excluding the unused ring position.
    {attribute 'OPC.UA.DA.Access' := '1'}
    BufferLength : UINT; //! Physical ring length; usable capacity is BufferLength minus one.
END_STRUCT
END_TYPE

// ---- Framework/EventBuffer/DataTypes/E_EventPublishResult.TcDUT
{region 'Documentation'}
(*!
<summary>Named non-positive event publishing results; positive INT results indicate successful insertion.</summary>
*)
{endregion}
{attribute 'qualified_only'}
TYPE E_EventPublishResult : E_FifoResult;
END_TYPE

// ---- Framework/EventBuffer/DataTypes/E_EventReservationResult.TcDUT
{region 'Documentation'}
(*!
<summary>Outcome of an immediate owner event-budget reservation.</summary>
*)
{endregion}
{attribute 'qualified_only'}
{attribute 'strict'}
TYPE E_EventReservationResult :
(
    Error := 0, //! Invalid prerequisite or permanently impossible budget; do not retry as capacity waiting.
    Accepted := 1, //! Owner and global reservation counts now reflect the requested budget.
    WaitingForCapacity := 2 //! Temporarily insufficient free capacity; counts unchanged and retry is allowed.
);
END_TYPE

// ---- Framework/EventBuffer/DataTypes/E_EventSeverity.TcDUT
{region 'Documentation'}
(*!
<summary>Logging severity, independent of test result.</summary>
*)
{endregion}
{attribute 'qualified_only'}
{attribute 'strict'}
TYPE E_EventSeverity :
(
    Trace := 0, //! Fine-grained execution tracing.
    Debug := 1, //! Diagnostic detail for investigation.
    Info := 2, //! Normal informational event.
    Warning := 3, //! Recoverable or noteworthy abnormal condition.
    Error := 4, //! An error diagnostic; does not itself define the owner's Result.
    Critical := 5 //! Critical diagnostic severity.
) USINT := Trace;
END_TYPE

// ---- Framework/EventBuffer/DataTypes/E_EventType.TcDUT
{region 'Documentation'}
(*!
<summary>Event payload classification.</summary>
*)
{endregion}
{attribute 'qualified_only'}
{attribute 'strict'}
TYPE E_EventType :
(
    Unknown := 0, //! No defined payload category.
    Result := 10, //! Owner or Assertion evaluation outcome.
    Trigger := 20, //! Lifecycle command accepted or reported by the owner.
    StateTransition := 30, //! Owner lifecycle transition.
    Info := 40, //! Informational event.
    Aggregation := 50, //! Owner counters and duration encoded for final aggregation.
    Framework := 60 //! Framework diagnostic rather than a test verdict.
) USINT := Unknown;
END_TYPE

// ---- Framework/EventBuffer/DataTypes/E_OwnerScope.TcDUT
{region 'Documentation'}
(*!
<summary>Semantic owner or technical diagnostic scope of an event.</summary>
*)
{endregion}
{attribute 'qualified_only'}
{attribute 'strict'}
TYPE E_OwnerScope :
(
    Unknown := 0, //! No defined owner category.
    Framework := 5, //! Framework-wide technical diagnostic.
    // SA0027: Qualified enum member; retained despite the analyzer's name-collision report.
    {attribute 'analysis' := '-27'}
    RunControl := 10, //! Root Run Control owner.
    TestSuiteOrchestrator := 15, //! Technical Suite-scheduling scope retained for event compatibility.
    TestSuite := 20, //! Test Suite owner.
    TestCaseOrchestrator := 25, //! Technical Test-Case-scheduling scope retained for event compatibility.
    TestCase := 30, //! Test Case owner.
    Assertion := 40, //! Assertion finding.
    Preparation := 50 //! Preparation diagnostic.
) USINT := Unknown;
END_TYPE

// ---- Framework/EventBuffer/DataTypes/ST_Event.TcDUT
{region 'Documentation'}
(*!
<summary>Event payload. Timestamp is UTC Unix nanoseconds; text is ASCII.</summary>
<description>
Constructors return unpublished values with SequenceId and Timestamp zero. The publisher assigns both; SequenceId alone governs order and acknowledgements. Nonzero loss makes the log incomplete. StateTransition records its destination; Framework diagnostics may record the related existing state instead.
</description>
*)
{endregion}
TYPE ST_Event :
STRUCT
    {attribute 'OPC.UA.DA.Access' := '1'}
    SequenceId : UDINT := 0; //! Producer-assigned event sequence within the current buffer epoch; zero is not a published event.
    {attribute 'OPC.UA.DA.Access' := '1'}
    Timestamp : LINT := 0; //! UTC Unix timestamp in nanoseconds, assigned on publication.
    {attribute 'OPC.UA.DA.Access' := '1'}
    OwnerScope : E_OwnerScope := E_OwnerScope.Unknown; //! Semantic owner or technical diagnostic scope; independent of the event type.
    {attribute 'OPC.UA.DA.Access' := '1'}
    EventType : E_EventType := E_EventType.Unknown; //! Payload category used by the consumer to interpret this event.
    {attribute 'OPC.UA.DA.Access' := '1'}
    Severity : E_EventSeverity := E_EventSeverity.Info; //! Logging severity, independent of Result.
    {attribute 'OPC.UA.DA.Access' := '1'}
    Name : STRING(GVL_Constants.NameLength) := ''; //! Hierarchical ASCII owner identity within NameLength.
    {attribute 'OPC.UA.DA.Access' := '1'}
    ResourceName : STRING(GVL_Constants.ResourceNameLength) := ''; //! Optional ASCII resource context; empty when not supplied.
    {attribute 'OPC.UA.DA.Access' := '1'}
    State : E_State := E_State.Uninitialized; //! Owner state associated with the event; transitions record their destination.
    {attribute 'OPC.UA.DA.Access' := '1'}
    Result : E_Result := E_Result.NotEvaluated; //! Evaluation result associated with the event; numeric order is not severity order.
    {attribute 'OPC.UA.DA.Access' := '1'}
    Message : STRING(GVL_Constants.MessageLength) := ''; //! ASCII diagnostic or category-specific payload text within MessageLength.
END_STRUCT
END_TYPE

// ---- Framework/EventBuffer/DataTypes/ST_EventBufferCommand.TcDUT
{region 'Documentation'}
(*!
<summary>External Event Buffer requests; zero sequence means no delete request.</summary>
<description>
Run Control handles Reset before Delete, attempts hierarchical reservation release and clears both commands after destructive reset. Delete clearing follows a captured-value comparison; a cleared request alone does not confirm deletion. Replacing a pending Delete request is permitted only with a higher valid contiguous watermark.
</description>
*)
{endregion}
TYPE ST_EventBufferCommand :
STRUCT
    {attribute 'OPC.UA.DA.Access' := '3'}
    Reset : BOOL := FALSE; //! Destructive buffer reset request; Run Control attempts subtree reservation release first and then clears this flag.
    {attribute 'OPC.UA.DA.Access' := '3'}
    DeleteSequenceId : UDINT := 0; //! Inclusive contiguous acknowledgement watermark; zero means no request. The buffer clears an unchanged request.
END_STRUCT
END_TYPE

// ---- Framework/EventBuffer/DataTypes/ST_EventBufferStatus.TcDUT
{region 'Documentation'}
(*!
<summary>Producer sequence, contiguous deletion watermark and loss count.</summary>
<description>
Sequence may advance before insertion succeeds, so gaps and a latest assigned value above the highest readable event are possible. The sequence saturates at UDINT maximum; reaching exhaustion is unsupported. LostEventCount saturates at UINT maximum and any nonzero count invalidates event-log completeness. Reset starts a new epoch with all three fields zero.
</description>
*)
{endregion}
TYPE ST_EventBufferStatus :
STRUCT
    {attribute 'OPC.UA.DA.Access' := '1'}
    SequenceId : UDINT := 0; //! Latest producer sequence in the current epoch, including attempted insertions.
    {attribute 'OPC.UA.DA.Access' := '1'}
    DeletedSequenceId : UDINT := 0; //! SequenceId of the last event actually released in the current epoch; request clearing alone is not deletion.
    {attribute 'OPC.UA.DA.Access' := '1'}
    LostEventCount : UINT := 0; //! Number of failed event insertions; saturates at UINT maximum until buffer reset.
END_STRUCT
END_TYPE

// ---- Framework/EventBuffer/DataTypes/ST_EventStream.TcDUT
{region 'Documentation'}
(*!
<summary>External Event Stream storage and producer-owned communication snapshots.</summary>
<description>
The array is actual producer-owned ring storage, not a periodically copied event view. Consumers validate ContractInfo, derive readable positions from FifoControl and use its BufferLength as the effective upper index. Only the separate Buffer command boundary is consumer-writable; reservation accounting is private.
</description>
*)
{endregion}
TYPE ST_EventStream :
STRUCT
    {attribute 'OPC.UA.DA.Access' := '1'}
    ContractInfo : ST_ContractInfo; //! Event-stream compatibility and framework version metadata.
    {attribute 'OPC.UA.DA.Access' := '1'}
    FifoControl : ST_FifoStatus := (ConfigError := TRUE); //! Producer-maintained ring indices, occupancy and validity snapshot.
    {attribute 'OPC.UA.DA.Access' := '1'}
    Status : ST_EventBufferStatus; //! Producer-maintained sequence, deletion watermark and loss snapshot.
    {attribute 'OPC.UA.DA.Access' := '1'}
    Buffer : ARRAY[1..Param_EventBuffer.EventBufferLength] OF ST_Event; //! Physical ring positions; one position remains unused.
END_STRUCT
END_TYPE

// ---- Framework/Preparation/DataTypes/ST_PreparationStatus.TcDUT
{region 'Documentation'}
(*!
<summary>Preparation progress; Ready does not imply Completed.</summary>
<description>
State is diagnostic progress of the Preparation, not the owning Test Case's lifecycle. Ready and Completed are independent observations. The concrete Preparation maintains a current consistent snapshot on every call, including disabled observation; querying Status does not refresh it or perform resource actions. Initial Unknown/Uninitialized values describe a not-yet-observed instance.
</description>
*)
{endregion}
TYPE ST_PreparationStatus :
STRUCT
    {attribute 'OPC.UA.DA.Access' := '1'}
    State : E_State := E_State.Uninitialized; //! Concrete Preparation state; independent of the coarse ExecutionStatus.
    {attribute 'OPC.UA.DA.Access' := '1'}
    ExecutionStatus : E_ExecutionStatus := E_ExecutionStatus.Unknown; //! Current observed preparation condition; not a retained test result.
    {attribute 'OPC.UA.DA.Access' := '1'}
    Ready : BOOL := FALSE; //! Resource can be driven to the target condition; FALSE while Running. Does not mean target reached.
    {attribute 'OPC.UA.DA.Access' := '1'}
    Running : BOOL := FALSE; //! Preparation is actively driving the resource toward its target.
    {attribute 'OPC.UA.DA.Access' := '1'}
    Completed : BOOL := FALSE; //! Target condition is currently reached; not latched by the base.
    {attribute 'OPC.UA.DA.Access' := '1'}
    Error : BOOL := FALSE; //! Preparation cannot continue meaningfully.
END_STRUCT
END_TYPE

// ---- Framework/RunControl/DataTypes/ST_RunConfig.TcDUT
{region 'Documentation'}
(*!
<summary>Run timing configuration; timeouts must be positive, CompletionDelay may be zero.</summary>
<description>
Configure supplies these root-owned timing values before initialization validation; runtime commands do not override them. Execution includes capacity waiting, ResetTimeout bounds the complete hierarchical reset and AbortTimeout bounds controlled termination. CompletionDelay holds Completing after one-shot final Result/Aggregation publication; even zero delay completes on a later call.
</description>
*)
{endregion}
TYPE ST_RunConfig :
STRUCT
    Timeout : TIME := T#30s; //! Positive execution timeout, including child progress; TIME uses milliseconds.
    ResetTimeout : TIME := T#1s; //! Positive Reset timeout, including event-capacity waiting; TIME uses milliseconds.
    AbortTimeout : TIME := T#1s; //! Positive timeout for controlled abort completion; TIME uses milliseconds.
    CompletionDelay : TIME := T#100ms; //! Delay in Completing before final Completed transition; zero allowed, default T#100ms.
END_STRUCT
END_TYPE

// ---- Framework/RunControl/DataTypes/ST_RunControl.TcDUT
{region 'Documentation'}
(*!
<summary>External Run Control projection; owner execution state is held separately.</summary>
<description>
The command adapter processes Cmd before the concrete owner call; the owner processes BufferCmd first and projects only Name and Status last. Bind the actual shared storage rather than copying the whole structure back, which could overwrite asynchronous consumer requests. Lifecycle Reset, destructive Buffer Reset and full hierarchical initialization are separate operations.
</description>
*)
{endregion}
TYPE ST_RunControl :
STRUCT
    {attribute 'OPC.UA.DA.Access' := '1'}
    Name : STRING(GVL_Constants.NameLength) := ''; //! Run Control identity projected after cyclic processing; consumer read-only.
    {attribute 'OPC.UA.DA.Access' := '3'}
    Cmd : ST_Command; //! Consumer-writable lifecycle requests handled by the external command adapter.
    {attribute 'OPC.UA.DA.Access' := '3'}
    BufferCmd : ST_EventBufferCommand; //! Consumer-writable event-buffer reset and acknowledgement requests handled by Run Control.
    {attribute 'OPC.UA.DA.Access' := '1'}
    Status : ST_RunControlStatus; //! Run Control execution/result snapshot projected after cyclic processing; consumer read-only.
END_STRUCT
END_TYPE

// ---- Framework/RunControl/DataTypes/ST_RunControlCommunication.TcDUT
{region 'Documentation'}
(*!
<summary>Published Run Control metadata and external command/status data; no FB instance state.</summary>
<description>
This is the Direct Access publication below GVL_UnitTest.RunControl. Consumers validate its ContractInfo before interpreting data or writing Cmd/BufferCmd. The producer owns identity and status; only the declared command fields are externally writable. Current status is diagnostic/control data, not a replacement for missing event evidence.
</description>
*)
{endregion}
TYPE ST_RunControlCommunication :
STRUCT
    {attribute 'OPC.UA.DA.Access' := '1'}
    ContractInfo : ST_ContractInfo; //! Direct-access compatibility and framework version metadata.
    {attribute 'OPC.UA.DA.Access' := '3'}
    ControlData : ST_RunControl; //! Published command/status storage; only Cmd and BufferCmd are consumer-writable.
END_STRUCT
END_TYPE

// ---- Framework/RunControl/DataTypes/ST_RunControlStatus.TcDUT
{region 'Documentation'}
(*!
<summary>Aggregated child execution counts and elapsed owner duration.</summary>
<description>
Execution and result counters are different observations, not disjoint categories to sum. Child calls and counters continue after the root result and final event payload have been held. Runtime is the root's active execution interval, including waits, projected to saturating TIME milliseconds; it is not the sum of Suite durations or the completion delay.
</description>
*)
{endregion}
TYPE ST_RunControlStatus :
STRUCT
    {attribute 'OPC.UA.DA.Access' := '1'}
    Execution : ST_ExecutionStatus; //! Owner lifecycle, readiness, result and error snapshot.
    {attribute 'OPC.UA.DA.Access' := '1'}
    SuiteCountTotal : UINT := 0; //! Total number of Suites in the current collection.
    {attribute 'OPC.UA.DA.Access' := '1'}
    SuiteCountInactive : UINT := 0; //! Number of children observed inactive.
    {attribute 'OPC.UA.DA.Access' := '1'}
    SuiteCountIdle : UINT := 0; //! Number of children observed Idle.
    {attribute 'OPC.UA.DA.Access' := '1'}
    SuiteCountRunning : UINT := 0; //! Number of children observed running.
    {attribute 'OPC.UA.DA.Access' := '1'}
    SuiteCountCompleted : UINT := 0; //! Number of children observed completed, irrespective of outcome.
    {attribute 'OPC.UA.DA.Access' := '1'}
    SuiteCountPassed : UINT := 0; //! Number of Suites with Passed result.
    {attribute 'OPC.UA.DA.Access' := '1'}
    SuiteCountFailed : UINT := 0; //! Number of Suites with Failed result.
    {attribute 'OPC.UA.DA.Access' := '1'}
    SuiteCountError : UINT := 0; //! Number of Suites reporting an error.
    {attribute 'OPC.UA.DA.Access' := '1'}
    Runtime : TIME := T#0ms; //! Elapsed execution duration projected to TIME milliseconds; not a timeout configuration.
END_STRUCT
END_TYPE

// ---- Framework/RunControl/DataTypes/ST_TestSuiteCollectionConfig.TcDUT
{region 'Documentation'}
(*!
<summary>Finalized Suite collection bounds, population and orchestration configuration.</summary>
<description>
This is configuration metadata, not retained child storage. The occupied prefix starts at FirstIndex and contains Count entries; LastIndex includes unused capacity. Require IsValid before use and keep the actual array, children and slot assignments stable for execution. A new full initialization rebuilds the composition.
</description>
*)
{endregion}
TYPE ST_TestSuiteCollectionConfig :
STRUCT
    FirstIndex : DINT; //! Lower bound of the caller-owned child array; occupied entries start here.
    LastIndex : DINT; //! Upper bound of the complete child array, including unused capacity.
    Count : UINT; //! Number of registered children; occupied range is FirstIndex through FirstIndex + Count - 1.
    IsValid : BOOL; //! TRUE after successful finalization; FALSE configurations must not be used.
    Mode : E_OrchestrationMode; //! Scheduling strategy selected for this initialized collection.
END_STRUCT
END_TYPE

// ---- Framework/TestCases/DataTypes/ST_TestCaseConfig.TcDUT
{region 'Documentation'}
(*!
<summary>Test Case timeout configuration; identity is supplied separately during Initialize.</summary>
<description>
Copied by Initialize and held fixed for execution; every timeout must be positive. Timeout covers active Starting, Preparation and Test processing. PreparationTimeout bounds each active Preparation state and restarts on a permitted next-state transition. ResetTimeout begins on actual entry into Reset; parent reservation waiting happens before its Reset request and is supervised by the Suite. Abort escalation retains the original abort deadline.
</description>
*)
{endregion}
TYPE ST_TestCaseConfig :
STRUCT
    Timeout : TIME := T#5s; //! Positive execution timeout, including child progress; TIME uses milliseconds.
    PreparationTimeout : TIME := T#2s; //! Positive timeout per active Preparation state; TIME uses milliseconds.
    ResetTimeout : TIME := T#1s; //! Positive timeout from entry into Reset for scenario cleanup; TIME uses milliseconds.
    AbortTimeout : TIME := T#1s; //! Positive timeout for controlled abort completion; TIME uses milliseconds.
END_STRUCT
END_TYPE

// ---- Framework/TestCases/DataTypes/ST_TestCaseExecutionStatus.TcDUT
{region 'Documentation'}
(*!
<summary>Test Case execution snapshot including Preparation and Test activity.</summary>
<description>
This is a by-value lifecycle projection, not an external command or a separate state machine. Preparation and Test intervals both map to coarse Running with their respective activity flags. Completed does not mean Passed. Initial declaration defaults use Unknown; regular uninitialized projection uses NotReady and Uninitialized TRUE. The base does not use Inactive for selection.
</description>
*)
{endregion}
TYPE ST_TestCaseExecutionStatus :
STRUCT
    {attribute 'OPC.UA.DA.Access' := '1'}
    State : E_State := E_State.Uninitialized; //! Owner's detailed lifecycle state, including configured Test Case phases.
    {attribute 'OPC.UA.DA.Access' := '1'}
    ExecutionStatus : E_ExecutionStatus := E_ExecutionStatus.Unknown; //! Coarse execution classification derived from State.
    {attribute 'OPC.UA.DA.Access' := '1'}
    Result : E_Result := E_Result.NotEvaluated; //! Current held evaluation result; numeric order is not severity order.
    {attribute 'OPC.UA.DA.Access' := '1'}
    Uninitialized : BOOL := FALSE; //! TRUE while owner State is Uninitialized; successful Initialize alone does not complete the initial Reset.
    {attribute 'OPC.UA.DA.Access' := '1'}
    ConfigError : BOOL := FALSE; //! Owner setup is invalid or has not yet been validated.
    {attribute 'OPC.UA.DA.Access' := '1'}
    Ready : BOOL := FALSE; //! Owner is initialized, Idle and ready to accept Start.
    {attribute 'OPC.UA.DA.Access' := '1'}
    Running : BOOL := FALSE; //! Owner is in its active execution phase.
    {attribute 'OPC.UA.DA.Access' := '1'}
    Completed : BOOL := FALSE; //! Owner has reached its terminal Completed state; does not imply Passed.
    {attribute 'OPC.UA.DA.Access' := '1'}
    Aborted : BOOL := FALSE; //! Owner completed with Abort result.
    {attribute 'OPC.UA.DA.Access' := '1'}
    // SA0033: Contract status field retained even when not consumed by this application.
    {attribute 'analysis' := '-33'}
    Inactive : BOOL := FALSE; //! Contract-reserved inactive indication; retained for compatible consumers.
    {attribute 'OPC.UA.DA.Access' := '1'}
    Error : BOOL := FALSE; //! Owner reports an error, including Result = Error.
    {attribute 'OPC.UA.DA.Access' := '1'}
    PreparationActive : BOOL := FALSE; //! A configured Preparation state is currently active.
    {attribute 'OPC.UA.DA.Access' := '1'}
    TestActive : BOOL := FALSE; //! A configured Test state is currently active.
END_STRUCT
END_TYPE

// ---- Framework/TestCases/DataTypes/ST_TestCaseStatus.TcDUT
{region 'Documentation'}
(*!
<summary>Test Case status and lifecycle-capacity metadata.</summary>
<description>
Counts and lifecycle fields are refreshed during regular calls; Assertion results continue to be collected after Completed while the final owner result and emitted payload remain held. Total includes all contributed results, including NotEvaluated and Abort. State counts are validated projections: zero may also reflect an unset/invalid backing count; require successful initialization before using metadata for admission. Runtime is active owner duration in saturating TIME milliseconds, not summed child durations. External publication requires an explicit data wrapper, not owner instance symbols.
</description>
*)
{endregion}
TYPE ST_TestCaseStatus :
STRUCT
    {attribute 'OPC.UA.DA.Access' := '1'}
    Execution : ST_TestCaseExecutionStatus; //! Owner lifecycle, readiness, result and error snapshot.
    {attribute 'OPC.UA.DA.Access' := '1'}
    PreparationStateCount : UINT := 0; //! Configured number of Preparation states; zero means no Preparation phase.
    {attribute 'OPC.UA.DA.Access' := '1'}
    TestStateCount : UINT := 0; //! Configured number of Test states; at least one after successful initialization.
    {attribute 'OPC.UA.DA.Access' := '1'}
    AssertionCountTotal : UINT := 0; //! Total number of Assertion contributions in the current collection.
    {attribute 'OPC.UA.DA.Access' := '1'}
    AssertionCountPassed : UINT := 0; //! Number of Assertion contributions with Passed result.
    {attribute 'OPC.UA.DA.Access' := '1'}
    AssertionCountFailed : UINT := 0; //! Number of Assertion contributions with Failed result.
    {attribute 'OPC.UA.DA.Access' := '1'}
    AssertionCountError : UINT := 0; //! Number of Assertion contributions with Error result.
    {attribute 'OPC.UA.DA.Access' := '1'}
    Runtime : TIME := T#0ms; //! Elapsed execution duration projected to TIME milliseconds; not a timeout configuration.
END_STRUCT
END_TYPE

// ---- Framework/TestSuites/DataTypes/ST_TestCaseCollectionConfig.TcDUT
{region 'Documentation'}
(*!
<summary>Finalized collection bounds, population and orchestration configuration.</summary>
<description>
This is metadata, not child storage. The occupied prefix starts at FirstIndex and has Count entries; LastIndex includes unused capacity. Require IsValid before use and retain the actual array, child instances and slot assignments unchanged for execution. Full hierarchical initialization rebuilds the composition.
</description>
*)
{endregion}
TYPE ST_TestCaseCollectionConfig :
STRUCT
    FirstIndex : DINT; //! Lower bound of the caller-owned child array; occupied entries start here.
    LastIndex : DINT; //! Upper bound of the complete child array, including unused capacity.
    Count : UINT; //! Number of registered children; occupied range is FirstIndex through FirstIndex + Count - 1.
    IsValid : BOOL; //! TRUE after successful finalization; FALSE configurations must not be used.
    Mode : E_OrchestrationMode; //! Scheduling strategy selected for this initialized collection.
END_STRUCT
END_TYPE

// ---- Framework/TestSuites/DataTypes/ST_TestSuiteConfig.TcDUT
{region 'Documentation'}
(*!
<summary>One-shot Test Suite initialization values; all timeouts must be positive.</summary>
<description>
Copied during Initialize and held fixed through execution; all three limits are positive. Execution Timeout includes child progress and capacity waiting. ResetTimeout bounds active Suite Reset, including subordinate admission and cleanup; the root supervises waiting before dispatching this Suite's Reset. Abort escalation preserves its original deadline. Initialization is repeatable only through the coordinated startup path, not an active-run recovery command.
</description>
*)
{endregion}
TYPE ST_TestSuiteConfig :
STRUCT
    Timeout : TIME := T#10s; //! Positive execution timeout, including child progress; TIME uses milliseconds.
    ResetTimeout : TIME := T#1s; //! Positive Reset timeout, including event-capacity waiting; TIME uses milliseconds.
    AbortTimeout : TIME := T#1s; //! Positive timeout for controlled abort completion; TIME uses milliseconds.
END_STRUCT
END_TYPE

// ---- Framework/TestSuites/DataTypes/ST_TestSuiteStatus.TcDUT
{region 'Documentation'}
(*!
<summary>Aggregated child execution counts and elapsed owner duration.</summary>
<description>
Execution and result counters are different, overlapping observations rather than one partition. Child calls and counters continue after the final owner result and published aggregation are held. Runtime is owner active execution time projected to saturating TIME milliseconds, not summed child duration. The childless mock keeps all Test Case counters zero.
</description>
*)
{endregion}
TYPE ST_TestSuiteStatus :
STRUCT
    {attribute 'OPC.UA.DA.Access' := '1'}
    Execution : ST_ExecutionStatus; //! Owner lifecycle, readiness, result and error snapshot.
    {attribute 'OPC.UA.DA.Access' := '1'}
    TestCaseCountTotal : UINT := 0; //! Total number of Test Cases in the current collection.
    {attribute 'OPC.UA.DA.Access' := '1'}
    TestCaseCountInactive : UINT := 0; //! Number of children observed inactive.
    {attribute 'OPC.UA.DA.Access' := '1'}
    TestCaseCountIdle : UINT := 0; //! Number of children observed Idle.
    {attribute 'OPC.UA.DA.Access' := '1'}
    TestCaseCountRunning : UINT := 0; //! Number of children observed running.
    {attribute 'OPC.UA.DA.Access' := '1'}
    TestCaseCountCompleted : UINT := 0; //! Number of children observed completed, irrespective of outcome.
    {attribute 'OPC.UA.DA.Access' := '1'}
    TestCaseCountPassed : UINT := 0; //! Number of Test Cases with Passed result.
    {attribute 'OPC.UA.DA.Access' := '1'}
    TestCaseCountFailed : UINT := 0; //! Number of Test Cases with Failed result.
    {attribute 'OPC.UA.DA.Access' := '1'}
    TestCaseCountError : UINT := 0; //! Number of Test Cases reporting an error.
    {attribute 'OPC.UA.DA.Access' := '1'}
    Runtime : TIME := T#0ms; //! Elapsed execution duration projected to TIME milliseconds; not a timeout configuration.
END_STRUCT
END_TYPE

// ---- SelfTests/Helper/Orchestration/DataTypes/E_OrchestrationArrayLayout.TcDUT
{region 'Documentation'}
(*!
<summary>Selects an actual fixed array used by the collection-bound tests.</summary>
*)
{endregion}
{attribute 'qualified_only'}
{attribute 'strict'}
TYPE E_OrchestrationArrayLayout :
(
    Ordinary, //! One-based three-entry fixture array.
    Shifted, //! Fixture array with lower bound 7.
    Negative, //! Fixture array with lower bound -3.
    SpareCapacity //! Six-entry fixture array with an occupied prefix and unused capacity.
);
END_TYPE

// ---- SelfTests/Helper/Orchestration/DataTypes/ST_OrchestrationCalls.TcDUT
{region 'Documentation'}
(*!
<summary>Per-cycle child interface calls; resource release counts only nonempty contributions separately.</summary>
*)
{endregion}
TYPE ST_OrchestrationCalls :
STRUCT
    StartCount : UINT; //! Start requests received during this fixture cycle.
    ResetCount : UINT; //! Reset requests received during this fixture cycle.
    AbortCount : UINT; //! Abort requests received during this fixture cycle.
    ExecutionReservationCount : UINT; //! Execution admission attempts during this fixture cycle, including rejected attempts.
    ResetReservationCount : UINT; //! Reset admission attempts during this fixture cycle, including rejected attempts.
    FreeCount : UINT; //! Reservation-release calls during this fixture cycle, including repeated empty releases.
    ReleasedEntryCount : UINT; //! Sum of local reservation markers cleared during this fixture cycle.
    BodyCount : UINT; //! Concrete child-body calls during this fixture cycle.
    StartWithoutReservation : BOOL; //! TRUE if Start was requested without the local admission marker.
    ResetWithoutReservation : BOOL; //! TRUE if Reset was requested without the local admission marker.
END_STRUCT
END_TYPE

// ---- SelfTests/Helper/Orchestration/DataTypes/ST_OrchestrationCycle.TcDUT
{region 'Documentation'}
(*!
<summary>Retained evidence for one helper call followed by one call per registered child.</summary>
*)
{endregion}
TYPE ST_OrchestrationCycle :
STRUCT
    Calls : ARRAY[1..3] OF ST_OrchestrationCalls; //! Per-child interface-call trace for this fixture cycle.
    BeforeChildren : ARRAY[1..3] OF ST_OrchestrationObservation; //! Child views after helper execution and before concrete child-body calls.
    AfterChildren : ARRAY[1..3] OF ST_OrchestrationObservation; //! Child views after concrete child-body calls.
    Reservations : ARRAY[1..3] OF UINT; //! Per-child local admission markers after this cycle.
    ActiveSlot : UINT; //! Helper execution slot observed for this cycle.
    ExecutionFinished : BOOL; //! Helper execution-completion indication for this cycle.
    Result : E_Result; //! Helper technical result for this cycle.
    Ready : BOOL; //! Helper readiness indication for this cycle.
    Task : E_OrchestratorTask; //! Task assigned to the helper for this cycle.
    HelperDidNotCallChildren : BOOL; //! TRUE if helper execution left all concrete child-body counters unchanged.
    RequestsDidNotChangeState : BOOL; //! TRUE if helper requests left the child observations unchanged before their body calls.
    ActiveChildCount : UINT; //! Number of children requested to Start in this cycle or observed in Starting through Completing before their body calls.
    ResetFinished : BOOL; //! Helper Reset-completion indication for this cycle.
    AbortFinished : BOOL; //! Helper Abort-completion indication for this cycle.
    TaskComplete : BOOL; //! Helper completion indication for the assigned task.
    ResetActive : BOOL; //! Helper assigned-task indication for Reset.
    ExecutionActive : BOOL; //! Helper assigned-task indication for Execution.
    AbortActive : BOOL; //! Helper assigned-task indication for Abort.
END_STRUCT
END_TYPE

// ---- SelfTests/Helper/Orchestration/DataTypes/ST_OrchestrationObservation.TcDUT
{region 'Documentation'}
(*!
<summary>Scripted child view applied only by its FB call, after helper processing.</summary>
*)
{endregion}
TYPE ST_OrchestrationObservation :
STRUCT
    State : E_State := E_State.Idle; //! Child lifecycle state accepted by the next child-body call.
    Result : E_Result := E_Result.NotEvaluated; //! Child result accepted by the next child-body call.
    Ready : BOOL := TRUE; //! Scripted child readiness accepted by the next child-body call.
    Complete : BOOL; //! Scripted terminal completion accepted by the next child-body call.
END_STRUCT
END_TYPE

// ---- SelfTests/Helper/Orchestration/DataTypes/ST_OrchestrationStep.TcDUT
{region 'Documentation'}
(*!
<summary>Independent stimulus and expected observations for one helper-then-children cycle.</summary>
*)
{endregion}
TYPE ST_OrchestrationStep :
STRUCT
    Task : E_OrchestratorTask := E_OrchestratorTask.Execution; //! Helper task to execute at this scripted checkpoint.
    Children : ARRAY[1..3] OF ST_OrchestrationObservation; //! Scripted observations installed by the child calls after helper execution.
    ExecutionReservationResults : ARRAY[1..3] OF E_EventReservationResult := [3(E_EventReservationResult.Accepted)]; //! Reservation responses are installed before the helper call; child observations follow afterwards.
    ResetReservationResults : ARRAY[1..3] OF E_EventReservationResult := [3(E_EventReservationResult.Accepted)]; //! Per-child Reset admission responses installed before helper execution.
    ExpectedUnacceptedExecutionReservations : ARRAY[1..3] OF UINT; //! Additional attempts returning WaitingForCapacity or Error, without a corresponding request.
    ExpectedUnacceptedResetReservations : ARRAY[1..3] OF UINT; //! Expected additional Reset admission attempts returning WaitingForCapacity or Error without a Reset request.
    MaxActiveChildCount : UINT := 1; //! Upper bound on active children during Execution, including this cycle's Start; Serial defaults to one.
    ExpectedStartChild : UINT; //! One-based child position expected to receive Start; zero means none.
    ExpectedSlot : UINT; //! Expected helper execution slot after this cycle.
    ExpectedFinished : BOOL; //! Expected helper execution-completion indication.
    ExpectedReady : BOOL; //! Expected helper readiness indication.
    ExpectedReservations : ARRAY[1..3] OF UINT; //! Expected per-child local reservation markers after this cycle.
    ExpectedReleasedEntries : ARRAY[1..3] OF UINT; //! Expected per-child sum of released markers during this cycle.
    ExpectedResetChild : UINT; //! One-based child position expected to receive Reset; zero means none.
    ExpectedAbortRequests : ARRAY[1..3] OF UINT; //! Expected per-child Abort-request counts during this cycle.
    ExpectedResetFinished : BOOL; //! Expected helper Reset-completion indication.
    ExpectedAbortFinished : BOOL; //! Expected helper Abort-completion indication.
    ExpectedResult : E_Result := E_Result.NotEvaluated; //! Expected helper technical result.
    ExpectedDiagnosticCount : UDINT; //! Expected cumulative diagnostic publications in the retained isolated capture.
END_STRUCT
END_TYPE

// ---- SelfTests/TestCases/TestSuite_AssertionFloatingPoint/DataTypes/FloatingPointBits_LReal.TcDUT
{region 'Documentation'}
(*!
<summary>Selftest-only IEEE LREAL bit view; no numeric conversion or stored addresses.</summary>
*)
{endregion}
TYPE FloatingPointBits_LReal :
UNION
    Bits : LWORD; //! Raw IEEE binary64 bit view of the shared storage; no numeric conversion.
    Value : LREAL; //! 64-bit floating-point view of the same shared storage.
END_UNION
END_TYPE

// ---- SelfTests/TestCases/TestSuite_AssertionFloatingPoint/DataTypes/FloatingPointBits_Real.TcDUT
{region 'Documentation'}
(*!
<summary>Selftest-only IEEE REAL bit view; no numeric conversion or stored addresses.</summary>
*)
{endregion}
TYPE FloatingPointBits_Real :
UNION
    Bits : DWORD; //! Raw IEEE binary32 bit view of the shared storage; no numeric conversion.
    Value : REAL; //! 32-bit floating-point view of the same shared storage.
END_UNION
END_TYPE

// ---- SelfTests/TestCases/TestSuite_CommandAdapter/DataTypes/E_AdapterCommand.TcDUT
{region 'Documentation'}
(*!
<summary>Selects one external lifecycle command for isolated qualification tests.</summary>
*)
{endregion}
{attribute 'qualified_only'}
{attribute 'strict'}
TYPE E_AdapterCommand :
(
    Start, //! Exercise the external Start command.
    Abort, //! Exercise the external Abort command.
    Reset //! Exercise the external Reset command.
);
END_TYPE

// ---- SelfTests/TestCases/TestSuite_RunControlLifecycle/DataTypes/E_RunControlCompletionScenario.TcDUT
{region 'Documentation'}
(*!
<summary>Completion-delay and retained-publication scenarios for the isolated root.</summary>
*)
{endregion}
{attribute 'qualified_only'}
{attribute 'strict'}
TYPE E_RunControlCompletionScenario :
(
    ZeroDelay, //! Complete with zero configured completion delay.
    DefaultDelay, //! Complete after the configured default delay.
    InvalidTime, //! Force invalid completion-time validity through the protected seam.
    LateResetChildren //! Exercise delayed child Reset completion after owner finalization.
);
END_TYPE

// ---- SelfTests/TestCases/TestSuite_RunControlLifecycle/DataTypes/E_RunControlLifecycleScenario.TcDUT
{region 'Documentation'}
(*!
<summary>Root failure and Abort stimuli, including continued Reset and preserved Abort deadlines after an error.</summary>
*)
{endregion}
{attribute 'qualified_only'}
{attribute 'strict'}
TYPE E_RunControlLifecycleScenario :
(
    ResetError, //! Script helper Error during owner Reset.
    ResetTimeout, //! Hold child Reset completion beyond the configured deadline.
    ResetErrorTimeout, //! Combine Reset helper Error with held Reset completion.
    ChildError, //! Script a child technical Error during execution.
    UnexpectedChildAbort, //! Script an unexpected child abort during execution.
    ExecutionError, //! Script helper Error during execution.
    ExecutionTimeout, //! Hold execution completion beyond the configured deadline.
    Abort, //! Request normal owner Abort.
    AbortError, //! Script helper Error during Abort.
    AbortTimeout, //! Hold Abort completion beyond the configured deadline.
    AbortErrorTimeout //! Combine Abort helper Error with held Abort completion.
);
END_TYPE

// ---- SelfTests/TestCases/TestSuite_TestSuiteLifecycle/DataTypes/E_SuiteLifecycleScenario.TcDUT
{region 'Documentation'}
(*!
<summary>Distinct owner failure/Abort stimuli; each instance keeps its selected scenario for the complete run.</summary>
*)
{endregion}
{attribute 'qualified_only'}
{attribute 'strict'}
TYPE E_SuiteLifecycleScenario :
(
    ResetError, //! Script helper Error during owner Reset.
    ResetTimeout, //! Hold child Reset completion beyond the configured deadline.
    ChildError, //! Script a child technical Error during execution.
    UnexpectedChildAbort, //! Script an unexpected child abort during execution.
    ExecutionError, //! Script helper Error during execution.
    ExecutionTimeout, //! Hold execution completion beyond the configured deadline.
    Abort, //! Request normal owner Abort.
    AbortError, //! Script helper Error during Abort.
    AbortTimeout //! Hold Abort completion beyond the configured deadline.
);
END_TYPE

// ---- Framework/Assertions/GlobalVariables/Param_Assertions.TcGVL
{region 'Documentation'}
(*!
<summary>Consumer-configurable text capacities for string assertions.</summary>
*)
{endregion}
{attribute 'qualified_only'}
VAR_GLOBAL CONSTANT
    {attribute 'TcNoSymbol'}
    AssertionStringLength : UINT := 80; //! STRING capacity, independent of diagnostic preview length.
    {attribute 'TcNoSymbol'}
    AssertionWStringLength : UINT := 80; //! WSTRING capacity in characters, independent of diagnostic preview length.
END_VAR

// ---- Framework/Common/GlobalVariables/Global_Version.TcGVL
{attribute 'TcGenerated'}
{attribute 'no-analysis'}
{attribute 'linkalways'}
// This function has been automatically generated from the project information.
VAR_GLOBAL CONSTANT
	{attribute 'const_non_replaced'}
	stLibVersion_Tc3_UnitTest : ST_LibVersion := (iMajor := 1, iMinor := 0, iBuild := 0, iRevision := 0, nFlags := 0, sVersion := '1.0.0.0');
END_VAR

// ---- Framework/Common/GlobalVariables/GVL_Constants.TcGVL
{region 'Documentation'}
(*!
<summary>Fixed framework capacities, lifecycle event allowances and communication contract versions.</summary>
*)
{endregion}
{attribute 'qualified_only'}
VAR_GLOBAL CONSTANT
    {attribute 'TcNoSymbol'}
    NameLength : UINT := 80; //! Maximum ASCII owner-name content length, excluding the terminator; part of the event contract.

    {attribute 'TcNoSymbol'}
    ResourceNameLength : UINT := 32; //! Maximum ASCII resource-name content length, excluding the terminator.
    {attribute 'TcNoSymbol'}
    MessageLength : UINT := 254; //! Maximum ASCII event-message content length, excluding the terminator.
    {attribute 'TcNoSymbol'}
    AssertionValueLength : UINT := 40; //! Maximum diagnostic value-preview content length; independent of input text capacity.

    {attribute 'TcNoSymbol'}
    VersionLength : UINT := 10; //! Maximum version-text content length for Major.Minor.Build, excluding the terminator.
    {attribute 'TcNoSymbol'}
    DirectAccessContractVersion : STRING(VersionLength) := '1.0.0'; //! Version of the PLC-owned Run Control direct-access contract.
    {attribute 'TcNoSymbol'}
    EventStreamContractVersion : STRING(VersionLength) := '1.0.0'; //! Version of the PLC-owned event-stream transfer and acknowledgement contract.

    {attribute 'TcNoSymbol'}
    TestSuiteExecutionEventCount : UINT := 10; //! Own Suite lifecycle events only; child reservations remain independent.
    {attribute 'TcNoSymbol'}
    TestSuiteResetEventCount : UINT := 4; //! Own Suite Reset-event allowance in entries; child reservations remain independent.
    {attribute 'TcNoSymbol'}
    TestCaseResetEventCount : UINT := 3; //! Own Test Case Reset-event allowance in entries.
END_VAR

// ---- Framework/Common/GlobalVariables/GVL_UnitTest.TcGVL
{region 'Documentation'}
(*!
<summary>Library-owned PLC/PC communication storage; only command fields are consumer-writable.</summary>
*)
{endregion}
{attribute 'qualified_only'}
{attribute 'linkalways'}
VAR_GLOBAL
    {attribute 'OPC.UA.DA' := '1'}
    {attribute 'OPC.UA.DA.Access' := '3'}
    // SA0027: Qualified communication symbol; intentionally named independently of the concrete FB.
    {attribute 'analysis' := '-27'}
    RunControl : ST_RunControlCommunication := (ContractInfo := (
        ContractVersion := GVL_Constants.DirectAccessContractVersion,
        FrameworkVersion := GetFrameworkVersion())); //! Published lifecycle command/status storage; only command members are consumer-writable.

    {attribute 'OPC.UA.DA' := '1'}
    {attribute 'OPC.UA.DA.Access' := '1'}
    EventStream : ST_EventStream := (ContractInfo := (
        ContractVersion := GVL_Constants.EventStreamContractVersion,
        FrameworkVersion := GetFrameworkVersion())); //! Published producer-owned event data and metadata; consumers acknowledge through RunControl.ControlData.BufferCmd.
END_VAR

// ---- Framework/EventBuffer/GlobalVariables/GVL_EventBuffer.TcGVL
{region 'Documentation'}
(*!
<summary>Default PLC-side event service and publisher binding; communication storage is in GVL_UnitTest.</summary>
<description>
Instance needs explicit storage initialization; declaring the GVL does not initialize the service. Publisher initially references Instance. Keep replacement publisher instances alive for all users retaining that interface; a global rebinding does not promise to replace previously retained instance-local bindings.
</description>
*)
{endregion}
{attribute 'qualified_only'}
VAR_GLOBAL
    {attribute 'TcNoSymbol'}
    Instance : EventBuffer; //! Default library event-buffer service; its storage is supplied separately at startup.
    {attribute 'TcNoSymbol'}
    Publisher : I_EventPublisher := Instance; //! Default publisher view initially bound to Instance; instance-local publisher bindings may override it.
END_VAR

// ---- Framework/EventBuffer/GlobalVariables/Param_EventBuffer.TcGVL
{region 'Documentation'}
(*!
<summary>Consumer-configurable compile-time capacities; no runtime command storage.</summary>
<description>
Library parameter defaults are consumer-overridable at compile time. EventBufferLength must be 3..32767; effective usable capacity is length minus one. Reset and execution headroom remain shared unreserved producer capacity, not a budget multiplied by active owners. Owner admission validates its complete budget against actual publisher capacity. External consumers use the published BufferLength rather than a local parameter value.
</description>
*)
{endregion}
{attribute 'qualified_only'}
VAR_GLOBAL CONSTANT
    {attribute 'TcNoSymbol'}
    EventBufferLength : UINT := 256; //! Physical ring length 3..32767, default 256; usable capacity is length minus one.
    {attribute 'TcNoSymbol'}
    EventBufferResetHeadroom : UINT := 20; //! Shared free producer capacity during hierarchical reset; must fit the buffer.
    {attribute 'TcNoSymbol'}
    EventBufferExecutionHeadroom : UINT := 10; //! Shared unreserved producer capacity during normal execution; must fit the buffer.
END_VAR

// ---- Framework/Assertions/Interfaces/I_Assertion.TcIO
{region 'Documentation'}
(*!
<summary>Assertion-specific identity and result view; initialization remains an instance API.</summary>
*)
{endregion}
INTERFACE I_Assertion EXTENDS I_ResultProvider

END_INTERFACE

// ---- Framework/Common/Interfaces/I_Orchestratable.TcIO
{region 'Documentation'}
(*!
<summary>Common child orchestration view; the owner calls the concrete FB.</summary>
*)
{endregion}
INTERFACE I_Orchestratable EXTENDS I_ResultProvider

{region 'Documentation'}
(*!
<summary>Parent-assigned slot; set only during configuration. Initialize and Reset retain it.</summary>
*)
{endregion}
{attribute 'monitoring' := 'call'}
PROPERTY ExecutionSlot : UINT //! Parent-assigned slot; set only during configuration. Initialize and Reset retain it.
GET // PUBLIC
END_GET
SET // PUBLIC
END_SET
END_PROPERTY

{region 'Documentation'}
(*!
<summary>Releases the complete registered subtree synchronously without changing lifecycle states. Attempts all contributions; FALSE permits partial success. Repeated release is idempotent.</summary>
*)
{endregion}
METHOD FreeReservedEvents : BOOL //! TRUE when all subtree contributions were released; FALSE permits partial success.
END_METHOD

{region 'Documentation'}
(*!
<summary>Reports configuration or runtime error.</summary>
*)
{endregion}
{attribute 'monitoring' := 'call'}
PROPERTY HasError : BOOL //! Reports configuration or runtime error.
GET // PUBLIC
END_GET
END_PROPERTY

{region 'Documentation'}
(*!
<summary>Reports terminal lifecycle completion.</summary>
*)
{endregion}
{attribute 'monitoring' := 'call'}
PROPERTY IsComplete : BOOL //! Reports terminal lifecycle completion.
GET // PUBLIC
END_GET
END_PROPERTY

{region 'Documentation'}
(*!
<summary>Reports successful explicit initialization, not lifecycle readiness.</summary>
*)
{endregion}
{attribute 'monitoring' := 'call'}
PROPERTY IsInitialized : BOOL //! Reports successful explicit initialization, not lifecycle readiness.
GET // PUBLIC
END_GET
END_PROPERTY

{region 'Documentation'}
(*!
<summary>Reports current start readiness.</summary>
*)
{endregion}
{attribute 'monitoring' := 'call'}
PROPERTY IsReady : BOOL //! Reports current start readiness.
GET // PUBLIC
END_GET
END_PROPERTY

{region 'Documentation'}
(*!
<summary>Records an Abort request for cyclic processing.</summary>
*)
{endregion}
METHOD RequestAbort
END_METHOD

{region 'Documentation'}
(*!
<summary>Records a reset request for cyclic processing.</summary>
*)
{endregion}
METHOD RequestReset
END_METHOD

{region 'Documentation'}
(*!
<summary>Records a start request for cyclic processing.</summary>
*)
{endregion}
METHOD RequestStart
END_METHOD

{region 'Documentation'}
(*!
<summary>Own contribution to the global Event Buffer reservation; changed only with that aggregate.</summary>
*)
{endregion}
{attribute 'monitoring' := 'call'}
PROPERTY ReservedEntryCount : UINT //! Own contribution to the global Event Buffer reservation; changed only with that aggregate.
GET // PUBLIC
END_GET
END_PROPERTY

{region 'Documentation'}
(*!
<summary>Accepted updates the reservation; WaitingForCapacity is retryable, Error is not.</summary>
*)
{endregion}
METHOD ReserveExecutionEvents : E_EventReservationResult //! Accepted on success, WaitingForCapacity for retryable pressure, Error for invalid setup or an impossible budget.
END_METHOD

{region 'Documentation'}
(*!
<summary>Accepted updates the reservation; WaitingForCapacity is retryable, Error is not.</summary>
*)
{endregion}
METHOD ReserveResetEvents : E_EventReservationResult //! Accepted on success, WaitingForCapacity for retryable pressure, Error for invalid setup or an impossible budget.
END_METHOD

{region 'Documentation'}
(*!
<summary>Current owner lifecycle state.</summary>
*)
{endregion}
{attribute 'monitoring' := 'call'}
PROPERTY State : E_State //! Current owner lifecycle state.
GET // PUBLIC
END_GET
END_PROPERTY

END_INTERFACE

// ---- Framework/Common/Interfaces/I_OrchestratableCollection.TcIO
{region 'Documentation'}
(*!
<summary>Read-only indexed view of the registered, owner-held children.</summary>
<description>
The occupied prefix starts at ChildArrayLowerBound and contains ChildCount entries; ChildArrayUpperBound includes unused capacity. Before enabling regular execution, the owner validates this metadata and the nonzero initialized children. Keep bounds, population, child identities and slots fixed for execution; the scheduler caches the occupied bounds. Lookup uses the actual DINT array index, returns zero outside the occupied prefix and does not call a child FB.
</description>
*)
{endregion}
INTERFACE I_OrchestratableCollection

{region 'Documentation'}
(*!
<summary>Actual array lower bound; zero when no configuration is available.</summary>
*)
{endregion}
{attribute 'monitoring' := 'call'}
PROPERTY ChildArrayLowerBound : DINT //! Actual array lower bound; zero when no configuration is available.
GET // PUBLIC
END_GET
END_PROPERTY

{region 'Documentation'}
(*!
<summary>Actual array upper bound, including unused capacity; process only ChildCount entries.</summary>
*)
{endregion}
{attribute 'monitoring' := 'call'}
PROPERTY ChildArrayUpperBound : DINT //! Actual array upper bound, including unused capacity; process only ChildCount entries.
GET // PUBLIC
END_GET
END_PROPERTY

{region 'Documentation'}
(*!
<summary>Registered population starting at ChildArrayLowerBound; zero when unavailable.</summary>
*)
{endregion}
{attribute 'monitoring' := 'call'}
PROPERTY ChildCount : UINT //! Registered population starting at ChildArrayLowerBound; zero when unavailable.
GET // PUBLIC
END_GET
END_PROPERTY

{region 'Documentation'}
(*!
<summary>Returns the registered entry at its original array index; invalid access returns zero.</summary>
*)
{endregion}
METHOD GetChild : I_Orchestratable //! Registered child interface at Index; zero for an invalid or unoccupied index.
VAR_INPUT
    Index : DINT; //! Original child-array index, not a registration ordinal; valid children occupy LowerBound through LowerBound + Count - 1.
END_VAR
END_METHOD

END_INTERFACE

// ---- Framework/Common/Interfaces/I_Orchestrator.TcIO
{region 'Documentation'}
(*!
<summary>Owner-facing initialization, cyclic execution and observations of the selected scheduler.</summary>
<description>
Initialize with an owner-validated, nonempty, stable collection before Execute. The owner calls Execute once before all concrete child FBs in the same task; the helper dispatches requests, while the owner retains concrete calls, aggregation and timeout supervision. Do not execute the same helper both through Execute and its concrete FB body in one cycle.

The default Orchestrator admits at most one new Start or Reset per call; shared slots allow overlapping execution, not simultaneous admission. Repeating a task preserves progress, and completion never chooses the next task. Technical Error is held until Initialize or entry into a new Reset task; Idle does not clear it. Reset/Abort completion is separate from a successful outcome, so inspect Result as well as the corresponding completion flag.
</description>
*)
{endregion}
INTERFACE I_Orchestrator

{region 'Documentation'}
(*!
<summary>Last task supplied to the scheduler.</summary>
*)
{endregion}
{attribute 'monitoring' := 'call'}
PROPERTY CurrentTask : E_OrchestratorTask //! Last task supplied to the scheduler.
GET // PUBLIC
END_GET
END_PROPERTY

{region 'Documentation'}
(*!
<summary>Executes the selected task once, before the owner&#x27;s child FB calls.</summary>
*)
{endregion}
METHOD Execute
VAR_INPUT
    Task : E_OrchestratorTask; //! Owner-selected work for this call; a task change initializes its scheduling once.
END_VAR
END_METHOD

{region 'Documentation'}
(*!
<summary>Binds the validated collection and initializes scheduling before the first Execute call.</summary>
<description>
Capacity, occupied entries, naming and slots are owner/builder responsibilities. The owner must also accept child initialization before enabling regular execution. The default helper caches lower bound and count, not the capacity upper bound, and retains the collection interface for later indexed reads. A failed default initialization drops the old binding rather than preserving it as a fallback.
</description>
*)
{endregion}
METHOD Initialize : BOOL //! TRUE when the child collection is accepted and scheduling is initialized.
VAR_INPUT
    Collection : I_OrchestratableCollection; //! Initialized, stable child collection retained by the scheduler; its owner and children must outlive use.
    Name : STRING(GVL_Constants.NameLength); //! Hierarchical owner name used to identify events; must satisfy the naming contract.
    ResourceName : STRING(GVL_Constants.ResourceNameLength) := ''; //! Optional resource context for diagnostics; empty by default.
END_VAR
END_METHOD

{region 'Documentation'}
(*!
<summary>Current Abort task is finished, with reservations reconciled.</summary>
*)
{endregion}
{attribute 'monitoring' := 'call'}
PROPERTY IsAbortFinished : BOOL //! Current Abort task is finished, with reservations reconciled.
GET // PUBLIC
END_GET
END_PROPERTY

{region 'Documentation'}
(*!
<summary>Current Execution task completed all slots without a technical error.</summary>
*)
{endregion}
{attribute 'monitoring' := 'call'}
PROPERTY IsExecutionFinished : BOOL //! Current Execution task completed all slots without a technical error.
GET // PUBLIC
END_GET
END_PROPERTY

{region 'Documentation'}
(*!
<summary>Collection binding and occupied bounds were accepted by Initialize.</summary>
*)
{endregion}
{attribute 'monitoring' := 'call'}
PROPERTY IsInitialized : BOOL //! Collection binding and occupied bounds were accepted by Initialize.
GET // PUBLIC
END_GET
END_PROPERTY

{region 'Documentation'}
(*!
<summary>Execution may start from Idle with ready children, reconciled reservations and no held error.</summary>
*)
{endregion}
{attribute 'monitoring' := 'call'}
PROPERTY IsReady : BOOL //! Execution may start from Idle with ready children, reconciled reservations and no held error.
GET // PUBLIC
END_GET
END_PROPERTY

{region 'Documentation'}
(*!
<summary>Report whether Reset is the assigned task, including after completion until a task change.</summary>
*)
{endregion}
{attribute 'monitoring' := 'call'}
PROPERTY IsResetActive : BOOL //! TRUE while Reset is the assigned task; completion alone does not clear this indication.
GET // PUBLIC
END_GET
END_PROPERTY

{region 'Documentation'}
(*!
<summary>Current Reset task is finished; failed terminal children also count as finished.</summary>
*)
{endregion}
{attribute 'monitoring' := 'call'}
PROPERTY IsResetFinished : BOOL //! Current Reset task is finished; failed terminal children also count as finished.
GET // PUBLIC
END_GET
END_PROPERTY

